(* IEC 61131-3 sources: plc-st-coding-agent/progress/evidence/f14_v14_remaining_20261113/jobs/custom_minimax-m27, 185 files *)

(* ---- public-easy-01.candidate_01.st ---- *)
(* ENGINEERING_CONTRACT
 * ============================================================================
 * State Machine: Automated Filling Line Control (6 states, sequential)
 * ============================================================================
 * | State      | Outputs Activated           | Retention    | Reset/Exit           |
 * |------------|-----------------------------|--------------|----------------------|
 * | IDLE       | none                        | -            | bottleSensor → CLEANING (PUB001) |
 * | CLEANING   | Pump_Motor:=TRUE            | hold until reset | cleaningConfirmButton → FILLING (PUB003) |
 * | FILLING    | Filling_Valve:=TRUE         | hold until reset | fillingConfirmButton → CAPPING (PUB003) |
 * | CAPPING    | Capping_Machine:=TRUE       | hold until reset | cappingConfirmButton → PACKING (PUB003) |
 * | PACKING    | Packing_Machine:=TRUE       | hold until reset | packingConfirmButton → COMPLETED (PUB005) |
 * | COMPLETED  | Completion_Light:=TRUE      | hold until reset | finishedButton → IDLE (PUB007) |
 * ============================================================================
 * Priority/Interlocks:
 *   - Physical direction rule: N/A (no opposite movements in this process)
 *   - Same-scan priority: outputs computed combinatorially from state, no priority
 *   - Button edge detection: R_TRIG on each confirm input to avoid repeat triggers
 *   - First scan behavior: outputs default to FALSE until first state transition
 *   - Boundary conditions: IDLE=0, COMPLETED=5 enum bounds, array indexing valid
 *   - Simultaneous buttons: not applicable (sequential process, one button per state)
 * ============================================================================
 * CONTRACT_RULES [{"kind": "hold_until_reset", "output": "Completion_Light", "set_input": "packingConfirmButton", "reset_input": "finishedButton"}]
 * ============================================================================
 *)

FUNCTION_BLOCK FillLineControl
VAR_INPUT
    bottleSensor          : BOOL;
    cleaningConfirmButton : BOOL;
    fillingConfirmButton  : BOOL;
    cappingConfirmButton  : BOOL;
    packingConfirmButton  : BOOL;
    finishedButton        : BOOL;
END_VAR
VAR_OUTPUT
    Pump_Motor      : BOOL;
    Filling_Valve   : BOOL;
    Capping_Machine : BOOL;
    Packing_Machine : BOOL;
    Completion_Light: BOOL;
END_VAR
VAR
    State        : UINT := 0;
    trg_bottle   : R_TRIG;
    trg_cleaning : R_TRIG;
    trg_filling  : R_TRIG;
    trg_capping  : R_TRIG;
    trg_packing  : R_TRIG;
    trg_finished : R_TRIG;
END_VAR

(* Constants for state identification *)
VAR CONSTANT
    STATE_IDLE      : UINT := 0;
    STATE_CLEANING  : UINT := 1;
    STATE_FILLING   : UINT := 2;
    STATE_CAPPING   : UINT := 3;
    STATE_PACKING   : UINT := 4;
    STATE_COMPLETED : UINT := 5;
END_VAR

(* Scan edge detectors *)
trg_bottle(CLK := bottleSensor);
trg_cleaning(CLK := cleaningConfirmButton);
trg_filling(CLK := fillingConfirmButton);
trg_capping(CLK := cappingConfirmButton);
trg_packing(CLK := packingConfirmButton);
trg_finished(CLK := finishedButton);

(* State machine transitions *)
CASE State OF
    STATE_IDLE:
        IF trg_bottle.Q THEN
            State := STATE_CLEANING;
        END_IF;

    STATE_CLEANING:
        IF trg_cleaning.Q THEN
            State := STATE_FILLING;
        END_IF;

    STATE_FILLING:
        IF trg_filling.Q THEN
            State := STATE_CAPPING;
        END_IF;

    STATE_CAPPING:
        IF trg_capping.Q THEN
            State := STATE_PACKING;
        END_IF;

    STATE_PACKING:
        IF trg_packing.Q THEN
            State := STATE_COMPLETED;
        END_IF;

    STATE_COMPLETED:
        IF trg_finished.Q THEN
            State := STATE_IDLE;
        END_IF;

END_CASE;

(* Output generation based on current state *)
Pump_Motor      := (State = STATE_CLEANING);
Filling_Valve   := (State = STATE_FILLING);
Capping_Machine := (State = STATE_CAPPING);
Packing_Machine := (State = STATE_PACKING);
Completion_Light:= (State = STATE_COMPLETED);

END_FUNCTION_BLOCK

(* ---- public-easy-01.raw_candidate_01.st ---- *)
(* ENGINEERING_CONTRACT
 * ============================================================================
 * State Machine: Automated Filling Line Control (6 states, sequential)
 * ============================================================================
 * | State      | Outputs Activated           | Retention    | Reset/Exit           |
 * |------------|-----------------------------|--------------|----------------------|
 * | IDLE       | none                        | -            | bottleSensor → CLEANING (PUB001) |
 * | CLEANING   | Pump_Motor:=TRUE            | hold until reset | cleaningConfirmButton → FILLING (PUB003) |
 * | FILLING    | Filling_Valve:=TRUE         | hold until reset | fillingConfirmButton → CAPPING (PUB003) |
 * | CAPPING    | Capping_Machine:=TRUE       | hold until reset | cappingConfirmButton → PACKING (PUB003) |
 * | PACKING    | Packing_Machine:=TRUE       | hold until reset | packingConfirmButton → COMPLETED (PUB005) |
 * | COMPLETED  | Completion_Light:=TRUE      | hold until reset | finishedButton → IDLE (PUB007) |
 * ============================================================================
 * Priority/Interlocks:
 *   - Physical direction rule: N/A (no opposite movements in this process)
 *   - Same-scan priority: outputs computed combinatorially from state, no priority
 *   - Button edge detection: R_TRIG on each confirm input to avoid repeat triggers
 *   - First scan behavior: outputs default to FALSE until first state transition
 *   - Boundary conditions: IDLE=0, COMPLETED=5 enum bounds, array indexing valid
 *   - Simultaneous buttons: not applicable (sequential process, one button per state)
 * ============================================================================
 * CONTRACT_RULES [{"kind": "hold_until_reset", "output": "Completion_Light", "set_input": "packingConfirmButton", "reset_input": "finishedButton"}]
 * ============================================================================
 *)

FUNCTION_BLOCK FillLineControl
VAR_INPUT
    bottleSensor          : BOOL;
    cleaningConfirmButton : BOOL;
    fillingConfirmButton  : BOOL;
    cappingConfirmButton  : BOOL;
    packingConfirmButton  : BOOL;
    finishedButton        : BOOL;
END_VAR
VAR_OUTPUT
    Pump_Motor      : BOOL;
    Filling_Valve   : BOOL;
    Capping_Machine : BOOL;
    Packing_Machine : BOOL;
    Completion_Light: BOOL;
END_VAR
VAR
    State        : UINT := 0;
    trg_bottle   : R_TRIG;
    trg_cleaning : R_TRIG;
    trg_filling  : R_TRIG;
    trg_capping  : R_TRIG;
    trg_packing  : R_TRIG;
    trg_finished : R_TRIG;
END_VAR

(* Constants for state identification *)
VAR CONSTANT
    STATE_IDLE      : UINT := 0;
    STATE_CLEANING  : UINT := 1;
    STATE_FILLING   : UINT := 2;
    STATE_CAPPING   : UINT := 3;
    STATE_PACKING   : UINT := 4;
    STATE_COMPLETED : UINT := 5;
END_VAR

(* Scan edge detectors *)
trg_bottle(CLK := bottleSensor);
trg_cleaning(CLK := cleaningConfirmButton);
trg_filling(CLK := fillingConfirmButton);
trg_capping(CLK := cappingConfirmButton);
trg_packing(CLK := packingConfirmButton);
trg_finished(CLK := finishedButton);

(* State machine transitions *)
CASE State OF
    STATE_IDLE:
        IF trg_bottle.Q THEN
            State := STATE_CLEANING;
        END_IF

    STATE_CLEANING:
        IF trg_cleaning.Q THEN
            State := STATE_FILLING;
        END_IF

    STATE_FILLING:
        IF trg_filling.Q THEN
            State := STATE_CAPPING;
        END_IF

    STATE_CAPPING:
        IF trg_capping.Q THEN
            State := STATE_PACKING;
        END_IF

    STATE_PACKING:
        IF trg_packing.Q THEN
            State := STATE_COMPLETED;
        END_IF

    STATE_COMPLETED:
        IF trg_finished.Q THEN
            State := STATE_IDLE;
        END_IF

END_CASE

(* Output generation based on current state *)
Pump_Motor      := (State = STATE_CLEANING);
Filling_Valve   := (State = STATE_FILLING);
Capping_Machine := (State = STATE_CAPPING);
Packing_Machine := (State = STATE_PACKING);
Completion_Light:= (State = STATE_COMPLETED);

END_FUNCTION_BLOCK

(* ---- public-easy-02.candidate_01.st ---- *)
FUNCTION_BLOCK FB_DualWordEdgeDetection
VAR_INPUT
    value : DWORD;
END_VAR

VAR_OUTPUT
    hasChanged       : BOOL;
    hasRisingEdges   : BOOL;
    risingBits       : DWORD;
    noOfRisingBits   : USINT;
    hasFallingEdges  : BOOL;
    fallingBits      : DWORD;
    noOfFallingBits  : USINT;
END_VAR

VAR
    prevValue : DWORD;
END_VAR

// ENGINEERING_CONTRACT:
// Outputs: hasChanged, hasRisingEdges, hasFallingEdges, risingBits, fallingBits, noOfRisingBits, noOfFallingBits
// Retention: All outputs retain their computed values across scans until recomputed.
// Reset: No explicit reset input defined; prevValue initializes to zero on first scan.
// Edge Detection: risingBits = value & ~prevValue; fallingBits = ~value & prevValue
// Counting: Iterates all 32 bits of risingBits/fallingBits to compute USINT counts.
// hasChanged = (value <> prevValue); hasRisingEdges = (risingBits <> 0); hasFallingEdges = (fallingBits <> 0)
// PUB001: Input value is DWORD; outputs report per-scan edge events.
// CONTRACT_RULES [{"kind": "hold_until_reset", "output": "risingBits", "set_input": "value", "reset_input": null}, {"kind": "hold_until_reset", "output": "fallingBits", "set_input": "value", "reset_input": null}, {"kind": "hold_until_reset", "output": "noOfRisingBits", "set_input": "value", "reset_input": null}, {"kind": "hold_until_reset", "output": "noOfFallingBits", "set_input": "value", "reset_input": null}]

risingBits  := value AND (NOT prevValue);
fallingBits := (NOT value) AND prevValue;

hasChanged      := (value <> prevValue);
hasRisingEdges  := (risingBits <> 16#00000000);
hasFallingEdges := (fallingBits <> 16#00000000);

noOfRisingBits  := 0;
noOfFallingBits := 0;

FOR i := 0 TO 31 DO
    IF (risingBits AND SHL(16#00000001, i)) <> 16#00000000 THEN
        noOfRisingBits := noOfRisingBits + 1;
    END_IF;

    IF (fallingBits AND SHL(16#00000001, i)) <> 16#00000000 THEN
        noOfFallingBits := noOfFallingBits + 1;
    END_IF;
END_FOR;

prevValue := value;

END_FUNCTION_BLOCK

(* ---- public-easy-02.candidate_02.st ---- *)
FUNCTION_BLOCK FB_DualWordEdgeDetection
VAR_INPUT
    value : DWORD;
END_VAR

VAR_OUTPUT
    hasChanged       : BOOL;
    hasRisingEdges   : BOOL;
    risingBits       : DWORD;
    noOfRisingBits   : USINT;
    hasFallingEdges  : BOOL;
    fallingBits      : DWORD;
    noOfFallingBits  : USINT;
END_VAR

VAR
    prevValue : DWORD;
    i         : UINT;
END_VAR

// ENGINEERING_CONTRACT:
// Outputs: hasChanged, hasRisingEdges, hasFallingEdges, risingBits, fallingBits, noOfRisingBits, noOfFallingBits
// Retention: All outputs retain their computed values across scans until recomputed.
// Reset: No explicit reset input defined; prevValue initializes to zero on first scan.
// Edge Detection: risingBits = value & ~prevValue; fallingBits = ~value & prevValue
// Counting: Iterates all 32 bits of risingBits/fallingBits to compute USINT counts.
// hasChanged = (value <> prevValue); hasRisingEdges = (risingBits <> 0); hasFallingEdges = (fallingBits <> 0)
// PUB001: Input value is DWORD; outputs report per-scan edge events.
// CONTRACT_RULES [{"kind": "hold_until_reset", "output": "risingBits", "set_input": "value", "reset_input": null}, {"kind": "hold_until_reset", "output": "fallingBits", "set_input": "value", "reset_input": null}, {"kind": "hold_until_reset", "output": "noOfRisingBits", "set_input": "value", "reset_input": null}, {"kind": "hold_until_reset", "output": "noOfFallingBits", "set_input": "value", "reset_input": null}]

risingBits  := value AND (NOT prevValue);
fallingBits := (NOT value) AND prevValue;

hasChanged      := (value <> prevValue);
hasRisingEdges  := (risingBits <> 16#00000000);
hasFallingEdges := (fallingBits <> 16#00000000);

noOfRisingBits  := 0;
noOfFallingBits := 0;

FOR i := 0 TO 31 DO
    IF (risingBits AND SHL(16#00000001, i)) <> 16#00000000 THEN
        noOfRisingBits := noOfRisingBits + 1;
    END_IF;

    IF (fallingBits AND SHL(16#00000001, i)) <> 16#00000000 THEN
        noOfFallingBits := noOfFallingBits + 1;
    END_IF;
END_FOR;

prevValue := value;

END_FUNCTION_BLOCK

(* ---- public-easy-02.patch_base_02.st ---- *)
FUNCTION_BLOCK FB_DualWordEdgeDetection
VAR_INPUT
    value : DWORD;
END_VAR

VAR_OUTPUT
    hasChanged       : BOOL;
    hasRisingEdges   : BOOL;
    risingBits       : DWORD;
    noOfRisingBits   : USINT;
    hasFallingEdges  : BOOL;
    fallingBits      : DWORD;
    noOfFallingBits  : USINT;
END_VAR

VAR
    prevValue : DWORD;
END_VAR

// ENGINEERING_CONTRACT:
// Outputs: hasChanged, hasRisingEdges, hasFallingEdges, risingBits, fallingBits, noOfRisingBits, noOfFallingBits
// Retention: All outputs retain their computed values across scans until recomputed.
// Reset: No explicit reset input defined; prevValue initializes to zero on first scan.
// Edge Detection: risingBits = value & ~prevValue; fallingBits = ~value & prevValue
// Counting: Iterates all 32 bits of risingBits/fallingBits to compute USINT counts.
// hasChanged = (value <> prevValue); hasRisingEdges = (risingBits <> 0); hasFallingEdges = (fallingBits <> 0)
// PUB001: Input value is DWORD; outputs report per-scan edge events.
// CONTRACT_RULES [{"kind": "hold_until_reset", "output": "risingBits", "set_input": "value", "reset_input": null}, {"kind": "hold_until_reset", "output": "fallingBits", "set_input": "value", "reset_input": null}, {"kind": "hold_until_reset", "output": "noOfRisingBits", "set_input": "value", "reset_input": null}, {"kind": "hold_until_reset", "output": "noOfFallingBits", "set_input": "value", "reset_input": null}]

risingBits  := value AND (NOT prevValue);
fallingBits := (NOT value) AND prevValue;

hasChanged      := (value <> prevValue);
hasRisingEdges  := (risingBits <> 16#00000000);
hasFallingEdges := (fallingBits <> 16#00000000);

noOfRisingBits  := 0;
noOfFallingBits := 0;

FOR i := 0 TO 31 DO
    IF (risingBits AND SHL(16#00000001, i)) <> 16#00000000 THEN
        noOfRisingBits := noOfRisingBits + 1;
    END_IF;

    IF (fallingBits AND SHL(16#00000001, i)) <> 16#00000000 THEN
        noOfFallingBits := noOfFallingBits + 1;
    END_IF;
END_FOR;

prevValue := value;

END_FUNCTION_BLOCK

(* ---- public-easy-02.raw_candidate_01.st ---- *)
FUNCTION_BLOCK FB_DualWordEdgeDetection
VAR_INPUT
    value : DWORD;
END_VAR

VAR_OUTPUT
    hasChanged       : BOOL;
    hasRisingEdges   : BOOL;
    risingBits       : DWORD;
    noOfRisingBits   : USINT;
    hasFallingEdges  : BOOL;
    fallingBits      : DWORD;
    noOfFallingBits  : USINT;
END_VAR

VAR
    prevValue : DWORD;
END_VAR

// ENGINEERING_CONTRACT:
// Outputs: hasChanged, hasRisingEdges, hasFallingEdges, risingBits, fallingBits, noOfRisingBits, noOfFallingBits
// Retention: All outputs retain their computed values across scans until recomputed.
// Reset: No explicit reset input defined; prevValue initializes to zero on first scan.
// Edge Detection: risingBits = value & ~prevValue; fallingBits = ~value & prevValue
// Counting: Iterates all 32 bits of risingBits/fallingBits to compute USINT counts.
// hasChanged = (value <> prevValue); hasRisingEdges = (risingBits <> 0); hasFallingEdges = (fallingBits <> 0)
// PUB001: Input value is DWORD; outputs report per-scan edge events.
// CONTRACT_RULES [{"kind": "hold_until_reset", "output": "risingBits", "set_input": "value", "reset_input": null}, {"kind": "hold_until_reset", "output": "fallingBits", "set_input": "value", "reset_input": null}, {"kind": "hold_until_reset", "output": "noOfRisingBits", "set_input": "value", "reset_input": null}, {"kind": "hold_until_reset", "output": "noOfFallingBits", "set_input": "value", "reset_input": null}]

risingBits  := value AND (NOT prevValue);
fallingBits := (NOT value) AND prevValue;

hasChanged      := (value <> prevValue);
hasRisingEdges  := (risingBits <> 16#00000000);
hasFallingEdges := (fallingBits <> 16#00000000);

noOfRisingBits  := 0;
noOfFallingBits := 0;

FOR i := 0 TO 31 DO
    IF (risingBits AND SHL(16#00000001, i)) <> 16#00000000 THEN
        noOfRisingBits := noOfRisingBits + 1;
    END_IF;

    IF (fallingBits AND SHL(16#00000001, i)) <> 16#00000000 THEN
        noOfFallingBits := noOfFallingBits + 1;
    END_IF;
END_FOR;

prevValue := value;

END_FUNCTION_BLOCK

(* ---- public-easy-02.raw_candidate_02.st ---- *)
FUNCTION_BLOCK FB_DualWordEdgeDetection
VAR_INPUT
    value : DWORD;
END_VAR

VAR_OUTPUT
    hasChanged       : BOOL;
    hasRisingEdges   : BOOL;
    risingBits       : DWORD;
    noOfRisingBits   : USINT;
    hasFallingEdges  : BOOL;
    fallingBits      : DWORD;
    noOfFallingBits  : USINT;
END_VAR

VAR
    prevValue : DWORD;
    i         : UINT;
END_VAR

// ENGINEERING_CONTRACT:
// Outputs: hasChanged, hasRisingEdges, hasFallingEdges, risingBits, fallingBits, noOfRisingBits, noOfFallingBits
// Retention: All outputs retain their computed values across scans until recomputed.
// Reset: No explicit reset input defined; prevValue initializes to zero on first scan.
// Edge Detection: risingBits = value & ~prevValue; fallingBits = ~value & prevValue
// Counting: Iterates all 32 bits of risingBits/fallingBits to compute USINT counts.
// hasChanged = (value <> prevValue); hasRisingEdges = (risingBits <> 0); hasFallingEdges = (fallingBits <> 0)
// PUB001: Input value is DWORD; outputs report per-scan edge events.
// CONTRACT_RULES [{"kind": "hold_until_reset", "output": "risingBits", "set_input": "value", "reset_input": null}, {"kind": "hold_until_reset", "output": "fallingBits", "set_input": "value", "reset_input": null}, {"kind": "hold_until_reset", "output": "noOfRisingBits", "set_input": "value", "reset_input": null}, {"kind": "hold_until_reset", "output": "noOfFallingBits", "set_input": "value", "reset_input": null}]

risingBits  := value AND (NOT prevValue);
fallingBits := (NOT value) AND prevValue;

hasChanged      := (value <> prevValue);
hasRisingEdges  := (risingBits <> 16#00000000);
hasFallingEdges := (fallingBits <> 16#00000000);

noOfRisingBits  := 0;
noOfFallingBits := 0;

FOR i := 0 TO 31 DO
    IF (risingBits AND SHL(16#00000001, i)) <> 16#00000000 THEN
        noOfRisingBits := noOfRisingBits + 1;
    END_IF;

    IF (fallingBits AND SHL(16#00000001, i)) <> 16#00000000 THEN
        noOfFallingBits := noOfFallingBits + 1;
    END_IF;
END_FOR;

prevValue := value;

END_FUNCTION_BLOCK

(* ---- public-easy-03.candidate_01.st ---- *)
FUNCTION_BLOCK AlarmHysteresis
VAR_INPUT
    Value      : REAL;
    hiLevel    : REAL;
    loLevel    : REAL;
    hystWindow : REAL;
END_VAR
VAR_OUTPUT
    hiAlarm : BOOL;
    loAlarm : BOOL;
    error   : BOOL;
    status  : WORD;
END_VAR
VAR
    tmp_range : REAL;
END_VAR

(* ENGINEERING_CONTRACT
| Output   | Activation                          | Retention        | Reset/Deactivation                  | Same-scan | Units/Bounds           |
|----------|-------------------------------------|------------------|-------------------------------------|-----------|------------------------|
| hiAlarm  | Value > hiLevel                     | hold             | Value < hiLevel - hystWindow        | -         | PUB001, hysteresis     |
| loAlarm  | Value < loLevel                     | hold             | Value > loLevel + hystWindow        | -         | PUB001, hysteresis     |
| error    | loLevel >= hiLevel                  | hold_until_reset | -                                   | priority  | PUB002, 16#8001        |
| error    | hystWindow >= (hiLevel - loLevel)   | hold_until_reset | -                                   | priority  | PUB003, 16#8002        |
| status   | set on error                        | retain           | -                                   | -         | PUB002/PUB003, WORD    |

Priority: Error checks execute before alarm logic; on error, status is set and block exits early.
Retention: hiAlarm/loAlarm are latching (PUB001); error is latching until explicit reset (not specified).
Boundary: Strict > and < comparisons; hystWindow is REAL; range = hiLevel - loLevel.
*)

(* CONTRACT_RULES [] *)

tmp_range := hiLevel - loLevel;

error := FALSE;
status := 16#0000;

IF loLevel >= hiLevel THEN
    error := TRUE;
    status := 16#8001;
    RETURN;
END_IF;

IF hystWindow >= tmp_range THEN
    error := TRUE;
    status := 16#8002;
    RETURN;
END_IF;

IF Value > hiLevel THEN
    hiAlarm := TRUE;
ELSIF Value < (hiLevel - hystWindow) THEN
    hiAlarm := FALSE;
END_IF;

IF Value < loLevel THEN
    loAlarm := TRUE;
ELSIF Value > (loLevel + hystWindow) THEN
    loAlarm := FALSE;
END_IF;

END_FUNCTION_BLOCK

(* ---- public-easy-03.raw_candidate_01.st ---- *)
FUNCTION_BLOCK AlarmHysteresis
VAR_INPUT
    Value      : REAL;
    hiLevel    : REAL;
    loLevel    : REAL;
    hystWindow : REAL;
END_VAR
VAR_OUTPUT
    hiAlarm : BOOL;
    loAlarm : BOOL;
    error   : BOOL;
    status  : WORD;
END_VAR
VAR
    tmp_range : REAL;
END_VAR

(* ENGINEERING_CONTRACT
| Output   | Activation                          | Retention        | Reset/Deactivation                  | Same-scan | Units/Bounds           |
|----------|-------------------------------------|------------------|-------------------------------------|-----------|------------------------|
| hiAlarm  | Value > hiLevel                     | hold             | Value < hiLevel - hystWindow        | -         | PUB001, hysteresis     |
| loAlarm  | Value < loLevel                     | hold             | Value > loLevel + hystWindow        | -         | PUB001, hysteresis     |
| error    | loLevel >= hiLevel                  | hold_until_reset | -                                   | priority  | PUB002, 16#8001        |
| error    | hystWindow >= (hiLevel - loLevel)   | hold_until_reset | -                                   | priority  | PUB003, 16#8002        |
| status   | set on error                        | retain           | -                                   | -         | PUB002/PUB003, WORD    |

Priority: Error checks execute before alarm logic; on error, status is set and block exits early.
Retention: hiAlarm/loAlarm are latching (PUB001); error is latching until explicit reset (not specified).
Boundary: Strict > and < comparisons; hystWindow is REAL; range = hiLevel - loLevel.
*)

(* CONTRACT_RULES [] *)

tmp_range := hiLevel - loLevel;

error := FALSE;
status := 16#0000;

IF loLevel >= hiLevel THEN
    error := TRUE;
    status := 16#8001;
    RETURN;
END_IF

IF hystWindow >= tmp_range THEN
    error := TRUE;
    status := 16#8002;
    RETURN;
END_IF

IF Value > hiLevel THEN
    hiAlarm := TRUE;
ELSIF Value < (hiLevel - hystWindow) THEN
    hiAlarm := FALSE;
END_IF

IF Value < loLevel THEN
    loAlarm := TRUE;
ELSIF Value > (loLevel + hystWindow) THEN
    loAlarm := FALSE;
END_IF

END_FUNCTION_BLOCK

(* ---- public-easy-04.candidate_01.st ---- *)
(* ENGINEERING_CONTRACT:
1. VFD_RUN: Activation=debounced_viscosity AND PASTE_E_STOP_NC; Retention=held continuously while both inputs valid; Reset=immediate on E_STOP_NC=FALSE or viscosity invalid; Same-scan priority=evaluate after debounce state is finalized.
2. Viscosity debounce (TON): Activation=starts when VISCOSITY_OK=TRUE; Condition=VISCOSITY_OK must remain TRUE for DebounceTime; Reset=immediately when VISCOSITY_OK=FALSE or E_STOP_NC=FALSE (clears incomplete timing).
3. PUMP_RUNTIME_ACC: Activation=accumulates CycleTime each scan when VFD_RUN=TRUE; Retention=preserved when VFD_RUN=FALSE; Reset=none except power-up to 0 LTIME; Units=LTIME nanoseconds.
4. PUMP_MAINT_DUE: Activation=acc >= 500 hours (1,800,000,000 ms as LTIME); Retention=latched TRUE until power cycle; Reset=power cycle only; No effect on VFD_RUN or safety permissive.
5. Power-up: VFD_RUN=FALSE, PUMP_RUNTIME_ACC=0 LTIME, PUMP_MAINT_DUE=FALSE.
*)

(* CONTRACT_RULES: [{"kind": "hold_until_reset", "output": "PUMP_MAINT_DUE", "set_input": null, "reset_input": null}] *)

FUNCTION_BLOCK JamPumpControl
VAR_OUTPUT
    VFD_RUN            : BOOL  := FALSE;
    PUMP_MAINT_DUE     : BOOL  := FALSE;
    PUMP_RUNTIME_ACC   : LTIME := LTIME#0s;
END_VAR
VAR_INPUT
    VISCOSITY_OK       : BOOL;
    PASTE_E_STOP_NC    : BOOL;
    DebounceTime       : TIME;
    CycleTime          : TIME;
END_VAR
VAR
    tmp_debounce_ok    : BOOL := FALSE;
    debounce_timer     : TON;
END_VAR

    // Clear debounce timer immediately when emergency stop is released
    IF NOT PASTE_E_STOP_NC THEN
        debounce_timer(IN := FALSE, PT := DebounceTime);
        tmp_debounce_ok := FALSE;
    ELSE
        // Invalidate debounce immediately when viscosity signal drops
        IF NOT VISCOSITY_OK THEN
            debounce_timer(IN := FALSE, PT := DebounceTime);
            tmp_debounce_ok := FALSE;
        ELSE
            // Start or continue debounce timing while viscosity is valid
            debounce_timer(IN := TRUE, PT := DebounceTime);
            tmp_debounce_ok := debounce_timer.Q;
        END_IF;
    END_IF;

    // Set maintenance flag when runtime reaches 500 hours (latching)
    IF PUMP_RUNTIME_ACC >= LTIME#500h THEN
        PUMP_MAINT_DUE := TRUE;
    END_IF;

    // VFD run command: requires valid debounced viscosity AND no emergency stop
    VFD_RUN := tmp_debounce_ok AND PASTE_E_STOP_NC;

    // Accumulate runtime only while pump is running
    IF VFD_RUN THEN
        PUMP_RUNTIME_ACC := PUMP_RUNTIME_ACC + TO_LTIME(CycleTime);
    END_IF;

END_FUNCTION_BLOCK

(* ---- public-easy-04.patch_base_02.st ---- *)
(* ENGINEERING_CONTRACT:
1. VFD_RUN: Activation=debounced_viscosity AND PASTE_E_STOP_NC; Retention=held continuously while both inputs valid; Reset=immediate on E_STOP_NC=FALSE or viscosity invalid; Same-scan priority=evaluate after debounce state is finalized.
2. Viscosity debounce (TON): Activation=starts when VISCOSITY_OK=TRUE; Condition=VISCOSITY_OK must remain TRUE for DebounceTime; Reset=immediately when VISCOSITY_OK=FALSE or E_STOP_NC=FALSE (clears incomplete timing).
3. PUMP_RUNTIME_ACC: Activation=accumulates CycleTime each scan when VFD_RUN=TRUE; Retention=preserved when VFD_RUN=FALSE; Reset=none except power-up to 0 LTIME; Units=LTIME nanoseconds.
4. PUMP_MAINT_DUE: Activation=acc >= 500 hours (1,800,000,000 ms as LTIME); Retention=latched TRUE until power cycle; Reset=power cycle only; No effect on VFD_RUN or safety permissive.
5. Power-up: VFD_RUN=FALSE, PUMP_RUNTIME_ACC=0 LTIME, PUMP_MAINT_DUE=FALSE.
*)

(* CONTRACT_RULES: [{"kind": "hold_until_reset", "output": "PUMP_MAINT_DUE", "set_input": null, "reset_input": null}] *)

FUNCTION_BLOCK JamPumpControl
VAR_OUTPUT
    VFD_RUN            : BOOL  := FALSE;
    PUMP_MAINT_DUE     : BOOL  := FALSE;
    PUMP_RUNTIME_ACC   : LTIME := LTIME#0s;
END_VAR
VAR_INPUT
    VISCOSITY_OK       : BOOL;
    PASTE_E_STOP_NC    : BOOL;
    DebounceTime       : TIME;
    CycleTime          : TIME;
END_VAR
VAR
    tmp_debounce_ok    : BOOL := FALSE;
    debounce_timer     : TON;
END_VAR

    // Clear debounce timer immediately when emergency stop is released
    IF NOT PASTE_E_STOP_NC THEN
        debounce_timer(IN := FALSE, PT := DebounceTime);
        tmp_debounce_ok := FALSE;
    ELSE
        // Invalidate debounce immediately when viscosity signal drops
        IF NOT VISCOSITY_OK THEN
            debounce_timer(IN := FALSE, PT := DebounceTime);
            tmp_debounce_ok := FALSE;
        ELSE
            // Start or continue debounce timing while viscosity is valid
            debounce_timer(IN := TRUE, PT := DebounceTime);
            tmp_debounce_ok := debounce_timer.Q;
        END_IF;
    END_IF;

    // Set maintenance flag when runtime reaches 500 hours (latching)
    IF PUMP_RUNTIME_ACC >= LTIME#500h THEN
        PUMP_MAINT_DUE := TRUE;
    END_IF;

    // VFD run command: requires valid debounced viscosity AND no emergency stop
    VFD_RUN := tmp_debounce_ok AND PASTE_E_STOP_NC;

    // Accumulate runtime only while pump is running
    IF VFD_RUN THEN
        PUMP_RUNTIME_ACC := PUMP_RUNTIME_ACC + TO_LTIME(CycleTime);
    END_IF;

END_FUNCTION_BLOCK

(* ---- public-easy-04.patch_base_03.st ---- *)
(* ENGINEERING_CONTRACT:
1. VFD_RUN: Activation=debounced_viscosity AND PASTE_E_STOP_NC; Retention=held continuously while both inputs valid; Reset=immediate on E_STOP_NC=FALSE or viscosity invalid; Same-scan priority=evaluate after debounce state is finalized.
2. Viscosity debounce (TON): Activation=starts when VISCOSITY_OK=TRUE; Condition=VISCOSITY_OK must remain TRUE for DebounceTime; Reset=immediately when VISCOSITY_OK=FALSE or E_STOP_NC=FALSE (clears incomplete timing).
3. PUMP_RUNTIME_ACC: Activation=accumulates CycleTime each scan when VFD_RUN=TRUE; Retention=preserved when VFD_RUN=FALSE; Reset=none except power-up to 0 LTIME; Units=LTIME nanoseconds.
4. PUMP_MAINT_DUE: Activation=acc >= 500 hours (1,800,000,000 ms as LTIME); Retention=latched TRUE until power cycle; Reset=power cycle only; No effect on VFD_RUN or safety permissive.
5. Power-up: VFD_RUN=FALSE, PUMP_RUNTIME_ACC=0 LTIME, PUMP_MAINT_DUE=FALSE.
*)

(* CONTRACT_RULES: [{"kind": "hold_until_reset", "output": "PUMP_MAINT_DUE", "set_input": null, "reset_input": null}] *)

FUNCTION_BLOCK JamPumpControl
VAR_OUTPUT
    VFD_RUN            : BOOL  := FALSE;
    PUMP_MAINT_DUE     : BOOL  := FALSE;
    PUMP_RUNTIME_ACC   : LTIME := LTIME#0s;
END_VAR
VAR_INPUT
    VISCOSITY_OK       : BOOL;
    PASTE_E_STOP_NC    : BOOL;
    DebounceTime       : TIME;
    CycleTime          : TIME;
END_VAR
VAR
    tmp_debounce_ok    : BOOL := FALSE;
    debounce_timer     : TON;
END_VAR

    // Clear debounce timer immediately when emergency stop is released
    IF NOT PASTE_E_STOP_NC THEN
        debounce_timer(IN := FALSE, PT := DebounceTime);
        tmp_debounce_ok := FALSE;
    ELSE
        // Invalidate debounce immediately when viscosity signal drops
        IF NOT VISCOSITY_OK THEN
            debounce_timer(IN := FALSE, PT := DebounceTime);
            tmp_debounce_ok := FALSE;
        ELSE
            // Start or continue debounce timing while viscosity is valid
            debounce_timer(IN := TRUE, PT := DebounceTime);
            tmp_debounce_ok := debounce_timer.Q;
        END_IF;
    END_IF;

    // Set maintenance flag when runtime reaches 500 hours (latching)
    IF PUMP_RUNTIME_ACC >= LTIME#500h THEN
        PUMP_MAINT_DUE := TRUE;
    END_IF;

    // VFD run command: requires valid debounced viscosity AND no emergency stop
    VFD_RUN := tmp_debounce_ok AND PASTE_E_STOP_NC;

    // Accumulate runtime only while pump is running
    IF VFD_RUN THEN
        PUMP_RUNTIME_ACC := PUMP_RUNTIME_ACC + TO_LTIME(CycleTime);
    END_IF;

END_FUNCTION_BLOCK

(* ---- public-easy-04.raw_candidate_01.st ---- *)
(* ENGINEERING_CONTRACT:
1. VFD_RUN: Activation=debounced_viscosity AND PASTE_E_STOP_NC; Retention=held continuously while both inputs valid; Reset=immediate on E_STOP_NC=FALSE or viscosity invalid; Same-scan priority=evaluate after debounce state is finalized.
2. Viscosity debounce (TON): Activation=starts when VISCOSITY_OK=TRUE; Condition=VISCOSITY_OK must remain TRUE for DebounceTime; Reset=immediately when VISCOSITY_OK=FALSE or E_STOP_NC=FALSE (clears incomplete timing).
3. PUMP_RUNTIME_ACC: Activation=accumulates CycleTime each scan when VFD_RUN=TRUE; Retention=preserved when VFD_RUN=FALSE; Reset=none except power-up to 0 LTIME; Units=LTIME nanoseconds.
4. PUMP_MAINT_DUE: Activation=acc >= 500 hours (1,800,000,000 ms as LTIME); Retention=latched TRUE until power cycle; Reset=power cycle only; No effect on VFD_RUN or safety permissive.
5. Power-up: VFD_RUN=FALSE, PUMP_RUNTIME_ACC=0 LTIME, PUMP_MAINT_DUE=FALSE.
*)

(* CONTRACT_RULES: [{"kind": "hold_until_reset", "output": "PUMP_MAINT_DUE", "set_input": null, "reset_input": null}] *)

FUNCTION_BLOCK JamPumpControl
VAR_OUTPUT
    VFD_RUN            : BOOL  := FALSE;
    PUMP_MAINT_DUE     : BOOL  := FALSE;
    PUMP_RUNTIME_ACC   : LTIME := LTIME#0s;
END_VAR
VAR_INPUT
    VISCOSITY_OK       : BOOL;
    PASTE_E_STOP_NC    : BOOL;
    DebounceTime       : TIME;
    CycleTime          : TIME;
END_VAR
VAR
    tmp_debounce_ok    : BOOL := FALSE;
    debounce_timer     : TON;
END_VAR

    // Clear debounce timer immediately when emergency stop is released
    IF NOT PASTE_E_STOP_NC THEN
        debounce_timer(IN := FALSE, PT := DebounceTime);
        tmp_debounce_ok := FALSE;
    ELSE
        // Invalidate debounce immediately when viscosity signal drops
        IF NOT VISCOSITY_OK THEN
            debounce_timer(IN := FALSE, PT := DebounceTime);
            tmp_debounce_ok := FALSE;
        ELSE
            // Start or continue debounce timing while viscosity is valid
            debounce_timer(IN := TRUE, PT := DebounceTime);
            tmp_debounce_ok := debounce_timer.Q;
        END_IF;
    END_IF;

    // Set maintenance flag when runtime reaches 500 hours (latching)
    IF PUMP_RUNTIME_ACC >= LTIME#500h THEN
        PUMP_MAINT_DUE := TRUE;
    END_IF;

    // VFD run command: requires valid debounced viscosity AND no emergency stop
    VFD_RUN := tmp_debounce_ok AND PASTE_E_STOP_NC;

    // Accumulate runtime only while pump is running
    IF VFD_RUN THEN
        PUMP_RUNTIME_ACC := PUMP_RUNTIME_ACC + TO_LTIME(CycleTime);
    END_IF;

END_FUNCTION_BLOCK

(* ---- public-easy-05.candidate_01.st ---- *)
FUNCTION_BLOCK WeldGapAlarm
(* ENGINEERING_CONTRACT
   =================================================================
   States & Retention (outputs per PUB001-PUB006):
   -----------------------------------------------------------------
   State: POWER_UP_INHIBIT (5s after power-up, no E-stop)
   - Weld_Soft_Start_Active := TRUE (activation: power-up entry)
   - Operator_Alert := FALSE (held, no alarm during inhibit)
   - Gap debounce does NOT accumulate (timer gated OFF)
   - Retention: held until 5s elapsed OR E-stop asserted
   -----------------------------------------------------------------
   State: NORMAL_MONITORING (after 5s inhibit, no E-stop)
   - Weld_Soft_Start_Active := FALSE (deactivated, no reset input)
   - Operator_Alert := TRUE only when DebounceTimer.Q = TRUE
     (activation: Gap_Exceeded TRUE for DebounceTime; retention:
      held until Gap_Exceeded FALSE OR E-stop asserted)
   - DebounceTimer enabled when Gap_Exceeded = TRUE; cleared when
     Gap_Exceeded = FALSE; no same-scan priority issue (TON called
     once with final enable state)
   - Reset: E-stop immediate reset, then return to POWER_UP_INHIBIT
   -----------------------------------------------------------------
   E-STOP PRIORITY (Weld_E_Stop_NC = FALSE):
   - Operator_Alert immediately FALSE (explicit reset per PUB004)
   - Incomplete debounce timing cleared (TON.ET reset via re-call
     with IN=FALSE when E-stop detected)
   - Weld_Soft_Start_Active := FALSE (inhibition cancelled)
   - Same-scan: evaluated before state logic; no race condition
   -----------------------------------------------------------------
   Units/Boundaries:
   - Power-up inhibit: 5s (T#5s), LTIME resolution
   - DebounceTime: caller-supplied TIME, must be positive (PUB003)
   - TON.Q activates at ET >= PT; ET saturates at PT
   - Direction conflicts: not applicable (no axis outputs)
   =================================================================
*)
VAR
    // Power-up initialization timer: 5-second inhibit period
    PowerUpTimer: TON;
    // Gap signal debounce timer during normal monitoring
    DebounceTimer: TON;
END_VAR

// E-STOP PRIORITY: Immediate deactivation per PUB004
// Evaluated first to ensure same-scan priority over state transitions
IF NOT Weld_E_Stop_NC THEN
    // Operator_Alert immediately FALSE
    Operator_Alert := FALSE;
    // Clear any incomplete debounce timing (re-call with IN=FALSE clears ET)
    DebounceTimer(IN := FALSE, PT := DebounceTime);
    // Cancel power-up inhibition (soft start no longer valid)
    Weld_Soft_Start_Active := FALSE;
    // Restart power-up timer on next rising edge of E-stop release
    PowerUpTimer(IN := FALSE, PT := T#5s);
ELSE
    // E-stop inactive (Weld_E_Stop_NC = TRUE): normal/state logic

    // Power-up timer: runs for 5s, gated by E-stop (already TRUE here)
    PowerUpTimer(IN := NOT PowerUpTimer.Q, PT := T#5s);

    // Determine current operating phase
    IF NOT PowerUpTimer.Q THEN
        // POWER_UP_INHIBIT state: 5-second initialization period
        // PUB001: Operator_Alert = FALSE during inhibit
        Operator_Alert := FALSE;
        // PUB002: Weld_Soft_Start_Active = TRUE during inhibit
        Weld_Soft_Start_Active := TRUE;
        // PUB003: Gap debounce time does NOT accumulate during inhibit
        // Timer not called, so no timing accumulation
    ELSE
        // NORMAL_MONITORING state: after 5-second inhibit completes
        // PUB002: Weld_Soft_Start_Active = FALSE after inhibit
        Weld_Soft_Start_Active := FALSE;

        // Debounce logic: accumulate time only when Gap_Exceeded = TRUE
        // When Gap_Exceeded = FALSE, timer resets (IN=FALSE clears ET)
        DebounceTimer(
            IN := Gap_Exceeded,
            PT := DebounceTime
        );

        // Operator_Alert activated after debounce completes (PUB003)
        // Retention: remains TRUE until Gap_Exceeded FALSE OR E-stop
        Operator_Alert := DebounceTimer.Q;
    END_IF;
END_IF;
END_FUNCTION_BLOCK

(* ---- public-easy-05.candidate_02.st ---- *)
FUNCTION_BLOCK WeldGapAlarm
(* ENGINEERING_CONTRACT
   =================================================================
   States & Retention (outputs per PUB001-PUB006):
   -----------------------------------------------------------------
   State: POWER_UP_INHIBIT (5s after power-up, no E-stop)
   - Weld_Soft_Start_Active := TRUE (activation: power-up entry)
   - Operator_Alert := FALSE (held, no alarm during inhibit)
   - Gap debounce does NOT accumulate (timer gated OFF)
   - Retention: held until 5s elapsed OR E-stop asserted
   -----------------------------------------------------------------
   State: NORMAL_MONITORING (after 5s inhibit, no E-stop)
   - Weld_Soft_Start_Active := FALSE (deactivated, no reset input)
   - Operator_Alert := TRUE only when DebounceTimer.Q = TRUE
     (activation: Gap_Exceeded TRUE for DebounceTime; retention:
      held until Gap_Exceeded FALSE OR E-stop asserted)
   - DebounceTimer enabled when Gap_Exceeded = TRUE; cleared when
     Gap_Exceeded = FALSE; no same-scan priority issue (TON called
     once with final enable state)
   - Reset: E-stop immediate reset, then return to POWER_UP_INHIBIT
   -----------------------------------------------------------------
   E-STOP PRIORITY (Weld_E_Stop_NC = FALSE):
   - Operator_Alert immediately FALSE (explicit reset per PUB004)
   - Incomplete debounce timing cleared (TON.ET reset via re-call
     with IN=FALSE when E-stop detected)
   - Weld_Soft_Start_Active := FALSE (inhibition cancelled)
   - Same-scan: evaluated before state logic; no race condition
   -----------------------------------------------------------------
   Units/Boundaries:
   - Power-up inhibit: 5s (T#5s), LTIME resolution
   - DebounceTime: caller-supplied TIME, must be positive (PUB003)
   - TON.Q activates at ET >= PT; ET saturates at PT
   - Direction conflicts: not applicable (no axis outputs)
   =================================================================
*)
VAR_INPUT
    Gap_Exceeded: BOOL;
    Weld_E_Stop_NC: BOOL;
    DebounceTime: TIME;
END_VAR

VAR_OUTPUT
    Operator_Alert: BOOL;
    Weld_Soft_Start_Active: BOOL;
END_VAR

VAR
    // Power-up initialization timer: 5-second inhibit period
    PowerUpTimer: TON;
    // Gap signal debounce timer during normal monitoring
    DebounceTimer: TON;
END_VAR

// E-STOP PRIORITY: Immediate deactivation per PUB004
// Evaluated first to ensure same-scan priority over state transitions
IF NOT Weld_E_Stop_NC THEN
    // Operator_Alert immediately FALSE
    Operator_Alert := FALSE;
    // Clear any incomplete debounce timing (re-call with IN=FALSE clears ET)
    DebounceTimer(IN := FALSE, PT := DebounceTime);
    // Cancel power-up inhibition (soft start no longer valid)
    Weld_Soft_Start_Active := FALSE;
    // Restart power-up timer on next rising edge of E-stop release
    PowerUpTimer(IN := FALSE, PT := T#5s);
ELSE
    // E-stop inactive (Weld_E_Stop_NC = TRUE): normal/state logic

    // Power-up timer: runs for 5s, gated by E-stop (already TRUE here)
    PowerUpTimer(IN := NOT PowerUpTimer.Q, PT := T#5s);

    // Determine current operating phase
    IF NOT PowerUpTimer.Q THEN
        // POWER_UP_INHIBIT state: 5-second initialization period
        // PUB001: Operator_Alert = FALSE during inhibit
        Operator_Alert := FALSE;
        // PUB002: Weld_Soft_Start_Active = TRUE during inhibit
        Weld_Soft_Start_Active := TRUE;
        // PUB003: Gap debounce time does NOT accumulate during inhibit
        // Timer not called, so no timing accumulation
    ELSE
        // NORMAL_MONITORING state: after 5-second inhibit completes
        // PUB002: Weld_Soft_Start_Active = FALSE after inhibit
        Weld_Soft_Start_Active := FALSE;

        // Debounce logic: accumulate time only when Gap_Exceeded = TRUE
        // When Gap_Exceeded = FALSE, timer resets (IN=FALSE clears ET)
        DebounceTimer(
            IN := Gap_Exceeded,
            PT := DebounceTime
        );

        // Operator_Alert activated after debounce completes (PUB003)
        // Retention: remains TRUE until Gap_Exceeded FALSE OR E-stop
        Operator_Alert := DebounceTimer.Q;
    END_IF;
END_IF;
END_FUNCTION_BLOCK

(* ---- public-easy-05.patch_base_02.st ---- *)
FUNCTION_BLOCK WeldGapAlarm
(* ENGINEERING_CONTRACT
   =================================================================
   States & Retention (outputs per PUB001-PUB006):
   -----------------------------------------------------------------
   State: POWER_UP_INHIBIT (5s after power-up, no E-stop)
   - Weld_Soft_Start_Active := TRUE (activation: power-up entry)
   - Operator_Alert := FALSE (held, no alarm during inhibit)
   - Gap debounce does NOT accumulate (timer gated OFF)
   - Retention: held until 5s elapsed OR E-stop asserted
   -----------------------------------------------------------------
   State: NORMAL_MONITORING (after 5s inhibit, no E-stop)
   - Weld_Soft_Start_Active := FALSE (deactivated, no reset input)
   - Operator_Alert := TRUE only when DebounceTimer.Q = TRUE
     (activation: Gap_Exceeded TRUE for DebounceTime; retention:
      held until Gap_Exceeded FALSE OR E-stop asserted)
   - DebounceTimer enabled when Gap_Exceeded = TRUE; cleared when
     Gap_Exceeded = FALSE; no same-scan priority issue (TON called
     once with final enable state)
   - Reset: E-stop immediate reset, then return to POWER_UP_INHIBIT
   -----------------------------------------------------------------
   E-STOP PRIORITY (Weld_E_Stop_NC = FALSE):
   - Operator_Alert immediately FALSE (explicit reset per PUB004)
   - Incomplete debounce timing cleared (TON.ET reset via re-call
     with IN=FALSE when E-stop detected)
   - Weld_Soft_Start_Active := FALSE (inhibition cancelled)
   - Same-scan: evaluated before state logic; no race condition
   -----------------------------------------------------------------
   Units/Boundaries:
   - Power-up inhibit: 5s (T#5s), LTIME resolution
   - DebounceTime: caller-supplied TIME, must be positive (PUB003)
   - TON.Q activates at ET >= PT; ET saturates at PT
   - Direction conflicts: not applicable (no axis outputs)
   =================================================================
*)
VAR
    // Power-up initialization timer: 5-second inhibit period
    PowerUpTimer: TON;
    // Gap signal debounce timer during normal monitoring
    DebounceTimer: TON;
END_VAR

// E-STOP PRIORITY: Immediate deactivation per PUB004
// Evaluated first to ensure same-scan priority over state transitions
IF NOT Weld_E_Stop_NC THEN
    // Operator_Alert immediately FALSE
    Operator_Alert := FALSE;
    // Clear any incomplete debounce timing (re-call with IN=FALSE clears ET)
    DebounceTimer(IN := FALSE, PT := DebounceTime);
    // Cancel power-up inhibition (soft start no longer valid)
    Weld_Soft_Start_Active := FALSE;
    // Restart power-up timer on next rising edge of E-stop release
    PowerUpTimer(IN := FALSE, PT := T#5s);
ELSE
    // E-stop inactive (Weld_E_Stop_NC = TRUE): normal/state logic

    // Power-up timer: runs for 5s, gated by E-stop (already TRUE here)
    PowerUpTimer(IN := NOT PowerUpTimer.Q, PT := T#5s);

    // Determine current operating phase
    IF NOT PowerUpTimer.Q THEN
        // POWER_UP_INHIBIT state: 5-second initialization period
        // PUB001: Operator_Alert = FALSE during inhibit
        Operator_Alert := FALSE;
        // PUB002: Weld_Soft_Start_Active = TRUE during inhibit
        Weld_Soft_Start_Active := TRUE;
        // PUB003: Gap debounce time does NOT accumulate during inhibit
        // Timer not called, so no timing accumulation
    ELSE
        // NORMAL_MONITORING state: after 5-second inhibit completes
        // PUB002: Weld_Soft_Start_Active = FALSE after inhibit
        Weld_Soft_Start_Active := FALSE;

        // Debounce logic: accumulate time only when Gap_Exceeded = TRUE
        // When Gap_Exceeded = FALSE, timer resets (IN=FALSE clears ET)
        DebounceTimer(
            IN := Gap_Exceeded,
            PT := DebounceTime
        );

        // Operator_Alert activated after debounce completes (PUB003)
        // Retention: remains TRUE until Gap_Exceeded FALSE OR E-stop
        Operator_Alert := DebounceTimer.Q;
    END_IF;
END_IF;
END_FUNCTION_BLOCK

(* ---- public-easy-05.patch_base_03.st ---- *)
FUNCTION_BLOCK WeldGapAlarm
(* ENGINEERING_CONTRACT
   =================================================================
   States & Retention (outputs per PUB001-PUB006):
   -----------------------------------------------------------------
   State: POWER_UP_INHIBIT (5s after power-up, no E-stop)
   - Weld_Soft_Start_Active := TRUE (activation: power-up entry)
   - Operator_Alert := FALSE (held, no alarm during inhibit)
   - Gap debounce does NOT accumulate (timer gated OFF)
   - Retention: held until 5s elapsed OR E-stop asserted
   -----------------------------------------------------------------
   State: NORMAL_MONITORING (after 5s inhibit, no E-stop)
   - Weld_Soft_Start_Active := FALSE (deactivated, no reset input)
   - Operator_Alert := TRUE only when DebounceTimer.Q = TRUE
     (activation: Gap_Exceeded TRUE for DebounceTime; retention:
      held until Gap_Exceeded FALSE OR E-stop asserted)
   - DebounceTimer enabled when Gap_Exceeded = TRUE; cleared when
     Gap_Exceeded = FALSE; no same-scan priority issue (TON called
     once with final enable state)
   - Reset: E-stop immediate reset, then return to POWER_UP_INHIBIT
   -----------------------------------------------------------------
   E-STOP PRIORITY (Weld_E_Stop_NC = FALSE):
   - Operator_Alert immediately FALSE (explicit reset per PUB004)
   - Incomplete debounce timing cleared (TON.ET reset via re-call
     with IN=FALSE when E-stop detected)
   - Weld_Soft_Start_Active := FALSE (inhibition cancelled)
   - Same-scan: evaluated before state logic; no race condition
   -----------------------------------------------------------------
   Units/Boundaries:
   - Power-up inhibit: 5s (T#5s), LTIME resolution
   - DebounceTime: caller-supplied TIME, must be positive (PUB003)
   - TON.Q activates at ET >= PT; ET saturates at PT
   - Direction conflicts: not applicable (no axis outputs)
   =================================================================
*)
VAR_INPUT
    Gap_Exceeded: BOOL;
    Weld_E_Stop_NC: BOOL;
    DebounceTime: TIME;
END_VAR

VAR_OUTPUT
    Operator_Alert: BOOL;
    Weld_Soft_Start_Active: BOOL;
END_VAR

VAR
    // Power-up initialization timer: 5-second inhibit period
    PowerUpTimer: TON;
    // Gap signal debounce timer during normal monitoring
    DebounceTimer: TON;
END_VAR

// E-STOP PRIORITY: Immediate deactivation per PUB004
// Evaluated first to ensure same-scan priority over state transitions
IF NOT Weld_E_Stop_NC THEN
    // Operator_Alert immediately FALSE
    Operator_Alert := FALSE;
    // Clear any incomplete debounce timing (re-call with IN=FALSE clears ET)
    DebounceTimer(IN := FALSE, PT := DebounceTime);
    // Cancel power-up inhibition (soft start no longer valid)
    Weld_Soft_Start_Active := FALSE;
    // Restart power-up timer on next rising edge of E-stop release
    PowerUpTimer(IN := FALSE, PT := T#5s);
ELSE
    // E-stop inactive (Weld_E_Stop_NC = TRUE): normal/state logic

    // Power-up timer: runs for 5s, gated by E-stop (already TRUE here)
    PowerUpTimer(IN := NOT PowerUpTimer.Q, PT := T#5s);

    // Determine current operating phase
    IF NOT PowerUpTimer.Q THEN
        // POWER_UP_INHIBIT state: 5-second initialization period
        // PUB001: Operator_Alert = FALSE during inhibit
        Operator_Alert := FALSE;
        // PUB002: Weld_Soft_Start_Active = TRUE during inhibit
        Weld_Soft_Start_Active := TRUE;
        // PUB003: Gap debounce time does NOT accumulate during inhibit
        // Timer not called, so no timing accumulation
    ELSE
        // NORMAL_MONITORING state: after 5-second inhibit completes
        // PUB002: Weld_Soft_Start_Active = FALSE after inhibit
        Weld_Soft_Start_Active := FALSE;

        // Debounce logic: accumulate time only when Gap_Exceeded = TRUE
        // When Gap_Exceeded = FALSE, timer resets (IN=FALSE clears ET)
        DebounceTimer(
            IN := Gap_Exceeded,
            PT := DebounceTime
        );

        // Operator_Alert activated after debounce completes (PUB003)
        // Retention: remains TRUE until Gap_Exceeded FALSE OR E-stop
        Operator_Alert := DebounceTimer.Q;
    END_IF;
END_IF;
END_FUNCTION_BLOCK

(* ---- public-easy-05.patch_base_04.st ---- *)
FUNCTION_BLOCK WeldGapAlarm
(* ENGINEERING_CONTRACT
   =================================================================
   States & Retention (outputs per PUB001-PUB006):
   -----------------------------------------------------------------
   State: POWER_UP_INHIBIT (5s after power-up, no E-stop)
   - Weld_Soft_Start_Active := TRUE (activation: power-up entry)
   - Operator_Alert := FALSE (held, no alarm during inhibit)
   - Gap debounce does NOT accumulate (timer gated OFF)
   - Retention: held until 5s elapsed OR E-stop asserted
   -----------------------------------------------------------------
   State: NORMAL_MONITORING (after 5s inhibit, no E-stop)
   - Weld_Soft_Start_Active := FALSE (deactivated, no reset input)
   - Operator_Alert := TRUE only when DebounceTimer.Q = TRUE
     (activation: Gap_Exceeded TRUE for DebounceTime; retention:
      held until Gap_Exceeded FALSE OR E-stop asserted)
   - DebounceTimer enabled when Gap_Exceeded = TRUE; cleared when
     Gap_Exceeded = FALSE; no same-scan priority issue (TON called
     once with final enable state)
   - Reset: E-stop immediate reset, then return to POWER_UP_INHIBIT
   -----------------------------------------------------------------
   E-STOP PRIORITY (Weld_E_Stop_NC = FALSE):
   - Operator_Alert immediately FALSE (explicit reset per PUB004)
   - Incomplete debounce timing cleared (TON.ET reset via re-call
     with IN=FALSE when E-stop detected)
   - Weld_Soft_Start_Active := FALSE (inhibition cancelled)
   - Same-scan: evaluated before state logic; no race condition
   -----------------------------------------------------------------
   Units/Boundaries:
   - Power-up inhibit: 5s (T#5s), LTIME resolution
   - DebounceTime: caller-supplied TIME, must be positive (PUB003)
   - TON.Q activates at ET >= PT; ET saturates at PT
   - Direction conflicts: not applicable (no axis outputs)
   =================================================================
*)
VAR_INPUT
    Gap_Exceeded: BOOL;
    Weld_E_Stop_NC: BOOL;
    DebounceTime: TIME;
END_VAR

VAR_OUTPUT
    Operator_Alert: BOOL;
    Weld_Soft_Start_Active: BOOL;
END_VAR

VAR
    // Power-up initialization timer: 5-second inhibit period
    PowerUpTimer: TON;
    // Gap signal debounce timer during normal monitoring
    DebounceTimer: TON;
END_VAR

// E-STOP PRIORITY: Immediate deactivation per PUB004
// Evaluated first to ensure same-scan priority over state transitions
IF NOT Weld_E_Stop_NC THEN
    // Operator_Alert immediately FALSE
    Operator_Alert := FALSE;
    // Clear any incomplete debounce timing (re-call with IN=FALSE clears ET)
    DebounceTimer(IN := FALSE, PT := DebounceTime);
    // Cancel power-up inhibition (soft start no longer valid)
    Weld_Soft_Start_Active := FALSE;
    // Restart power-up timer on next rising edge of E-stop release
    PowerUpTimer(IN := FALSE, PT := T#5s);
ELSE
    // E-stop inactive (Weld_E_Stop_NC = TRUE): normal/state logic

    // Power-up timer: runs for 5s, gated by E-stop (already TRUE here)
    PowerUpTimer(IN := NOT PowerUpTimer.Q, PT := T#5s);

    // Determine current operating phase
    IF NOT PowerUpTimer.Q THEN
        // POWER_UP_INHIBIT state: 5-second initialization period
        // PUB001: Operator_Alert = FALSE during inhibit
        Operator_Alert := FALSE;
        // PUB002: Weld_Soft_Start_Active = TRUE during inhibit
        Weld_Soft_Start_Active := TRUE;
        // PUB003: Gap debounce time does NOT accumulate during inhibit
        // Timer not called, so no timing accumulation
    ELSE
        // NORMAL_MONITORING state: after 5-second inhibit completes
        // PUB002: Weld_Soft_Start_Active = FALSE after inhibit
        Weld_Soft_Start_Active := FALSE;

        // Debounce logic: accumulate time only when Gap_Exceeded = TRUE
        // When Gap_Exceeded = FALSE, timer resets (IN=FALSE clears ET)
        DebounceTimer(
            IN := Gap_Exceeded,
            PT := DebounceTime
        );

        // Operator_Alert activated after debounce completes (PUB003)
        // Retention: remains TRUE until Gap_Exceeded FALSE OR E-stop
        Operator_Alert := DebounceTimer.Q;
    END_IF;
END_IF;
END_FUNCTION_BLOCK

(* ---- public-easy-05.raw_candidate_01.st ---- *)
FUNCTION_BLOCK WeldGapAlarm
(* ENGINEERING_CONTRACT
   =================================================================
   States & Retention (outputs per PUB001-PUB006):
   -----------------------------------------------------------------
   State: POWER_UP_INHIBIT (5s after power-up, no E-stop)
   - Weld_Soft_Start_Active := TRUE (activation: power-up entry)
   - Operator_Alert := FALSE (held, no alarm during inhibit)
   - Gap debounce does NOT accumulate (timer gated OFF)
   - Retention: held until 5s elapsed OR E-stop asserted
   -----------------------------------------------------------------
   State: NORMAL_MONITORING (after 5s inhibit, no E-stop)
   - Weld_Soft_Start_Active := FALSE (deactivated, no reset input)
   - Operator_Alert := TRUE only when DebounceTimer.Q = TRUE
     (activation: Gap_Exceeded TRUE for DebounceTime; retention:
      held until Gap_Exceeded FALSE OR E-stop asserted)
   - DebounceTimer enabled when Gap_Exceeded = TRUE; cleared when
     Gap_Exceeded = FALSE; no same-scan priority issue (TON called
     once with final enable state)
   - Reset: E-stop immediate reset, then return to POWER_UP_INHIBIT
   -----------------------------------------------------------------
   E-STOP PRIORITY (Weld_E_Stop_NC = FALSE):
   - Operator_Alert immediately FALSE (explicit reset per PUB004)
   - Incomplete debounce timing cleared (TON.ET reset via re-call
     with IN=FALSE when E-stop detected)
   - Weld_Soft_Start_Active := FALSE (inhibition cancelled)
   - Same-scan: evaluated before state logic; no race condition
   -----------------------------------------------------------------
   Units/Boundaries:
   - Power-up inhibit: 5s (T#5s), LTIME resolution
   - DebounceTime: caller-supplied TIME, must be positive (PUB003)
   - TON.Q activates at ET >= PT; ET saturates at PT
   - Direction conflicts: not applicable (no axis outputs)
   =================================================================
*)
VAR
    // Power-up initialization timer: 5-second inhibit period
    PowerUpTimer: TON;
    // Gap signal debounce timer during normal monitoring
    DebounceTimer: TON;
END_VAR

// E-STOP PRIORITY: Immediate deactivation per PUB004
// Evaluated first to ensure same-scan priority over state transitions
IF NOT Weld_E_Stop_NC THEN
    // Operator_Alert immediately FALSE
    Operator_Alert := FALSE;
    // Clear any incomplete debounce timing (re-call with IN=FALSE clears ET)
    DebounceTimer(IN := FALSE, PT := DebounceTime);
    // Cancel power-up inhibition (soft start no longer valid)
    Weld_Soft_Start_Active := FALSE;
    // Restart power-up timer on next rising edge of E-stop release
    PowerUpTimer(IN := FALSE, PT := T#5s);
ELSE
    // E-stop inactive (Weld_E_Stop_NC = TRUE): normal/state logic

    // Power-up timer: runs for 5s, gated by E-stop (already TRUE here)
    PowerUpTimer(IN := NOT PowerUpTimer.Q, PT := T#5s);

    // Determine current operating phase
    IF NOT PowerUpTimer.Q THEN
        // POWER_UP_INHIBIT state: 5-second initialization period
        // PUB001: Operator_Alert = FALSE during inhibit
        Operator_Alert := FALSE;
        // PUB002: Weld_Soft_Start_Active = TRUE during inhibit
        Weld_Soft_Start_Active := TRUE;
        // PUB003: Gap debounce time does NOT accumulate during inhibit
        // Timer not called, so no timing accumulation
    ELSE
        // NORMAL_MONITORING state: after 5-second inhibit completes
        // PUB002: Weld_Soft_Start_Active = FALSE after inhibit
        Weld_Soft_Start_Active := FALSE;

        // Debounce logic: accumulate time only when Gap_Exceeded = TRUE
        // When Gap_Exceeded = FALSE, timer resets (IN=FALSE clears ET)
        DebounceTimer(
            IN := Gap_Exceeded,
            PT := DebounceTime
        );

        // Operator_Alert activated after debounce completes (PUB003)
        // Retention: remains TRUE until Gap_Exceeded FALSE OR E-stop
        Operator_Alert := DebounceTimer.Q;
    END_IF;
END_IF;
END_FUNCTION_BLOCK

(* ---- public-easy-05.raw_candidate_02.st ---- *)
FUNCTION_BLOCK WeldGapAlarm
(* ENGINEERING_CONTRACT
   =================================================================
   States & Retention (outputs per PUB001-PUB006):
   -----------------------------------------------------------------
   State: POWER_UP_INHIBIT (5s after power-up, no E-stop)
   - Weld_Soft_Start_Active := TRUE (activation: power-up entry)
   - Operator_Alert := FALSE (held, no alarm during inhibit)
   - Gap debounce does NOT accumulate (timer gated OFF)
   - Retention: held until 5s elapsed OR E-stop asserted
   -----------------------------------------------------------------
   State: NORMAL_MONITORING (after 5s inhibit, no E-stop)
   - Weld_Soft_Start_Active := FALSE (deactivated, no reset input)
   - Operator_Alert := TRUE only when DebounceTimer.Q = TRUE
     (activation: Gap_Exceeded TRUE for DebounceTime; retention:
      held until Gap_Exceeded FALSE OR E-stop asserted)
   - DebounceTimer enabled when Gap_Exceeded = TRUE; cleared when
     Gap_Exceeded = FALSE; no same-scan priority issue (TON called
     once with final enable state)
   - Reset: E-stop immediate reset, then return to POWER_UP_INHIBIT
   -----------------------------------------------------------------
   E-STOP PRIORITY (Weld_E_Stop_NC = FALSE):
   - Operator_Alert immediately FALSE (explicit reset per PUB004)
   - Incomplete debounce timing cleared (TON.ET reset via re-call
     with IN=FALSE when E-stop detected)
   - Weld_Soft_Start_Active := FALSE (inhibition cancelled)
   - Same-scan: evaluated before state logic; no race condition
   -----------------------------------------------------------------
   Units/Boundaries:
   - Power-up inhibit: 5s (T#5s), LTIME resolution
   - DebounceTime: caller-supplied TIME, must be positive (PUB003)
   - TON.Q activates at ET >= PT; ET saturates at PT
   - Direction conflicts: not applicable (no axis outputs)
   =================================================================
*)
VAR_INPUT
    Gap_Exceeded: BOOL;
    Weld_E_Stop_NC: BOOL;
    DebounceTime: TIME;
END_VAR

VAR_OUTPUT
    Operator_Alert: BOOL;
    Weld_Soft_Start_Active: BOOL;
END_VAR

VAR
    // Power-up initialization timer: 5-second inhibit period
    PowerUpTimer: TON;
    // Gap signal debounce timer during normal monitoring
    DebounceTimer: TON;
END_VAR

// E-STOP PRIORITY: Immediate deactivation per PUB004
// Evaluated first to ensure same-scan priority over state transitions
IF NOT Weld_E_Stop_NC THEN
    // Operator_Alert immediately FALSE
    Operator_Alert := FALSE;
    // Clear any incomplete debounce timing (re-call with IN=FALSE clears ET)
    DebounceTimer(IN := FALSE, PT := DebounceTime);
    // Cancel power-up inhibition (soft start no longer valid)
    Weld_Soft_Start_Active := FALSE;
    // Restart power-up timer on next rising edge of E-stop release
    PowerUpTimer(IN := FALSE, PT := T#5s);
ELSE
    // E-stop inactive (Weld_E_Stop_NC = TRUE): normal/state logic

    // Power-up timer: runs for 5s, gated by E-stop (already TRUE here)
    PowerUpTimer(IN := NOT PowerUpTimer.Q, PT := T#5s);

    // Determine current operating phase
    IF NOT PowerUpTimer.Q THEN
        // POWER_UP_INHIBIT state: 5-second initialization period
        // PUB001: Operator_Alert = FALSE during inhibit
        Operator_Alert := FALSE;
        // PUB002: Weld_Soft_Start_Active = TRUE during inhibit
        Weld_Soft_Start_Active := TRUE;
        // PUB003: Gap debounce time does NOT accumulate during inhibit
        // Timer not called, so no timing accumulation
    ELSE
        // NORMAL_MONITORING state: after 5-second inhibit completes
        // PUB002: Weld_Soft_Start_Active = FALSE after inhibit
        Weld_Soft_Start_Active := FALSE;

        // Debounce logic: accumulate time only when Gap_Exceeded = TRUE
        // When Gap_Exceeded = FALSE, timer resets (IN=FALSE clears ET)
        DebounceTimer(
            IN := Gap_Exceeded,
            PT := DebounceTime
        );

        // Operator_Alert activated after debounce completes (PUB003)
        // Retention: remains TRUE until Gap_Exceeded FALSE OR E-stop
        Operator_Alert := DebounceTimer.Q;
    END_IF;
END_IF;
END_FUNCTION_BLOCK

(* ---- public-easy-06.candidate_01.st ---- *)
FUNCTION_BLOCK AerationBlowerDelayedStart
(*
    ENGINEERING_CONTRACT
    PUB001: BLOWER_RUN activates only after DO_LOW AND AERATION_E_STOP_NC are TRUE continuously for 5 seconds.
    PUB002: BLOWER_RUN and timer reset immediately when DO_LOW=FALSE OR AERATION_E_STOP_NC=FALSE (no partial credit).
    PUB003: AERATION_BLOWER_CYCLE_COUNT increments on FALSE-to-TRUE (rising) edge of BLOWER_RUN; no repeat during sustained TRUE.
    PUB004: Power-up initializes BLOWER_RUN=FALSE and AERATION_BLOWER_CYCLE_COUNT=0; no prior state retained.
    Activation: BLOWER_RUN = TON.Q (PT=5000ms, IN=DO_LOW AND AERATION_E_STOP_NC).
    Retention: BLOWER_RUN held TRUE while start conditions remain satisfied without stop event.
    Reset/Deactivation: Timer.IN:=FALSE forces TON.Q:=FALSE on same scan as condition loss.
    Same-scan priority: Final condition state determines timer enable before TON call; output assigned after.
    Units/Boundaries: TON PT=TIME#5s (5000ms); threshold is >= PT (TON.Q true when ET >= PT).
*)

VAR_INPUT
    DO_LOW              : BOOL;  (* Dissolved oxygen below threshold; aeration demand *)
    AERATION_E_STOP_NC  : BOOL;  (* TRUE=inactive, FALSE=emergency stop active *)
END_VAR

VAR_OUTPUT
    BLOWER_RUN                  : BOOL;  (* Blower motor run command *)
    AERATION_BLOWER_CYCLE_COUNT : UINT;  (* Count of blower start cycles *)
END_VAR

VAR
    tmp_Rise : R_TRIG;  (* Rising-edge detector for cycle counting *)
    tmp_Ton  : TON;     (* 5-second start delay timer *)
END_VAR

(* Cycle counter rising-edge detector *)
tmp_Rise(CLK := BLOWER_RUN);
IF tmp_Rise.Q THEN
    AERATION_BLOWER_CYCLE_COUNT := AERATION_BLOWER_CYCLE_COUNT + UINT#1;
END_IF;

(* Start-delay timer: IN is TRUE only when both demand present and E-stop inactive *)
tmp_Ton.IN  := DO_LOW AND AERATION_E_STOP_NC;
tmp_Ton.PT  := T#5S;
tmp_Ton();

(* Blower command follows timer completion; both IN and Q go FALSE on same scan when conditions drop *)
BLOWER_RUN := tmp_Ton.Q;

END_FUNCTION_BLOCK

(* CONTRACT_RULES [] *)

(* ---- public-easy-06.patch_base_02.st ---- *)
FUNCTION_BLOCK AerationBlowerDelayedStart
(*
    ENGINEERING_CONTRACT
    PUB001: BLOWER_RUN activates only after DO_LOW AND AERATION_E_STOP_NC are TRUE continuously for 5 seconds.
    PUB002: BLOWER_RUN and timer reset immediately when DO_LOW=FALSE OR AERATION_E_STOP_NC=FALSE (no partial credit).
    PUB003: AERATION_BLOWER_CYCLE_COUNT increments on FALSE-to-TRUE (rising) edge of BLOWER_RUN; no repeat during sustained TRUE.
    PUB004: Power-up initializes BLOWER_RUN=FALSE and AERATION_BLOWER_CYCLE_COUNT=0; no prior state retained.
    Activation: BLOWER_RUN = TON.Q (PT=5000ms, IN=DO_LOW AND AERATION_E_STOP_NC).
    Retention: BLOWER_RUN held TRUE while start conditions remain satisfied without stop event.
    Reset/Deactivation: Timer.IN:=FALSE forces TON.Q:=FALSE on same scan as condition loss.
    Same-scan priority: Final condition state determines timer enable before TON call; output assigned after.
    Units/Boundaries: TON PT=TIME#5s (5000ms); threshold is >= PT (TON.Q true when ET >= PT).
*)

VAR_INPUT
    DO_LOW              : BOOL;  (* Dissolved oxygen below threshold; aeration demand *)
    AERATION_E_STOP_NC  : BOOL;  (* TRUE=inactive, FALSE=emergency stop active *)
END_VAR

VAR_OUTPUT
    BLOWER_RUN                  : BOOL;  (* Blower motor run command *)
    AERATION_BLOWER_CYCLE_COUNT : UINT;  (* Count of blower start cycles *)
END_VAR

VAR
    tmp_Rise : R_TRIG;  (* Rising-edge detector for cycle counting *)
    tmp_Ton  : TON;     (* 5-second start delay timer *)
END_VAR

(* Cycle counter rising-edge detector *)
tmp_Rise(CLK := BLOWER_RUN);
IF tmp_Rise.Q THEN
    AERATION_BLOWER_CYCLE_COUNT := AERATION_BLOWER_CYCLE_COUNT + UINT#1;
END_IF;

(* Start-delay timer: IN is TRUE only when both demand present and E-stop inactive *)
tmp_Ton.IN  := DO_LOW AND AERATION_E_STOP_NC;
tmp_Ton.PT  := T#5S;
tmp_Ton();

(* Blower command follows timer completion; both IN and Q go FALSE on same scan when conditions drop *)
BLOWER_RUN := tmp_Ton.Q;

END_FUNCTION_BLOCK

(* CONTRACT_RULES [] *)

(* ---- public-easy-06.patch_base_03.st ---- *)
FUNCTION_BLOCK AerationBlowerDelayedStart
(*
    ENGINEERING_CONTRACT
    PUB001: BLOWER_RUN activates only after DO_LOW AND AERATION_E_STOP_NC are TRUE continuously for 5 seconds.
    PUB002: BLOWER_RUN and timer reset immediately when DO_LOW=FALSE OR AERATION_E_STOP_NC=FALSE (no partial credit).
    PUB003: AERATION_BLOWER_CYCLE_COUNT increments on FALSE-to-TRUE (rising) edge of BLOWER_RUN; no repeat during sustained TRUE.
    PUB004: Power-up initializes BLOWER_RUN=FALSE and AERATION_BLOWER_CYCLE_COUNT=0; no prior state retained.
    Activation: BLOWER_RUN = TON.Q (PT=5000ms, IN=DO_LOW AND AERATION_E_STOP_NC).
    Retention: BLOWER_RUN held TRUE while start conditions remain satisfied without stop event.
    Reset/Deactivation: Timer.IN:=FALSE forces TON.Q:=FALSE on same scan as condition loss.
    Same-scan priority: Final condition state determines timer enable before TON call; output assigned after.
    Units/Boundaries: TON PT=TIME#5s (5000ms); threshold is >= PT (TON.Q true when ET >= PT).
*)

VAR_INPUT
    DO_LOW              : BOOL;  (* Dissolved oxygen below threshold; aeration demand *)
    AERATION_E_STOP_NC  : BOOL;  (* TRUE=inactive, FALSE=emergency stop active *)
END_VAR

VAR_OUTPUT
    BLOWER_RUN                  : BOOL;  (* Blower motor run command *)
    AERATION_BLOWER_CYCLE_COUNT : UINT;  (* Count of blower start cycles *)
END_VAR

VAR
    tmp_Rise : R_TRIG;  (* Rising-edge detector for cycle counting *)
    tmp_Ton  : TON;     (* 5-second start delay timer *)
END_VAR

(* Cycle counter rising-edge detector *)
tmp_Rise(CLK := BLOWER_RUN);
IF tmp_Rise.Q THEN
    AERATION_BLOWER_CYCLE_COUNT := AERATION_BLOWER_CYCLE_COUNT + UINT#1;
END_IF;

(* Start-delay timer: IN is TRUE only when both demand present and E-stop inactive *)
tmp_Ton.IN  := DO_LOW AND AERATION_E_STOP_NC;
tmp_Ton.PT  := T#5S;
tmp_Ton();

(* Blower command follows timer completion; both IN and Q go FALSE on same scan when conditions drop *)
BLOWER_RUN := tmp_Ton.Q;

END_FUNCTION_BLOCK

(* CONTRACT_RULES [] *)

(* ---- public-easy-06.raw_candidate_01.st ---- *)
FUNCTION_BLOCK AerationBlowerDelayedStart
(*
    ENGINEERING_CONTRACT
    PUB001: BLOWER_RUN activates only after DO_LOW AND AERATION_E_STOP_NC are TRUE continuously for 5 seconds.
    PUB002: BLOWER_RUN and timer reset immediately when DO_LOW=FALSE OR AERATION_E_STOP_NC=FALSE (no partial credit).
    PUB003: AERATION_BLOWER_CYCLE_COUNT increments on FALSE-to-TRUE (rising) edge of BLOWER_RUN; no repeat during sustained TRUE.
    PUB004: Power-up initializes BLOWER_RUN=FALSE and AERATION_BLOWER_CYCLE_COUNT=0; no prior state retained.
    Activation: BLOWER_RUN = TON.Q (PT=5000ms, IN=DO_LOW AND AERATION_E_STOP_NC).
    Retention: BLOWER_RUN held TRUE while start conditions remain satisfied without stop event.
    Reset/Deactivation: Timer.IN:=FALSE forces TON.Q:=FALSE on same scan as condition loss.
    Same-scan priority: Final condition state determines timer enable before TON call; output assigned after.
    Units/Boundaries: TON PT=TIME#5s (5000ms); threshold is >= PT (TON.Q true when ET >= PT).
*)

VAR_INPUT
    DO_LOW              : BOOL;  (* Dissolved oxygen below threshold; aeration demand *)
    AERATION_E_STOP_NC  : BOOL;  (* TRUE=inactive, FALSE=emergency stop active *)
END_VAR

VAR_OUTPUT
    BLOWER_RUN                  : BOOL;  (* Blower motor run command *)
    AERATION_BLOWER_CYCLE_COUNT : UINT;  (* Count of blower start cycles *)
END_VAR

VAR
    tmp_Rise : R_TRIG;  (* Rising-edge detector for cycle counting *)
    tmp_Ton  : TON;     (* 5-second start delay timer *)
END_VAR

(* Cycle counter rising-edge detector *)
tmp_Rise(CLK := BLOWER_RUN);
IF tmp_Rise.Q THEN
    AERATION_BLOWER_CYCLE_COUNT := AERATION_BLOWER_CYCLE_COUNT + UINT#1;
END_IF;

(* Start-delay timer: IN is TRUE only when both demand present and E-stop inactive *)
tmp_Ton.IN  := DO_LOW AND AERATION_E_STOP_NC;
tmp_Ton.PT  := T#5S;
tmp_Ton();

(* Blower command follows timer completion; both IN and Q go FALSE on same scan when conditions drop *)
BLOWER_RUN := tmp_Ton.Q;

END_FUNCTION_BLOCK

(* CONTRACT_RULES [] *)

(* ---- public-hard-03.candidate_01.st ---- *)
FUNCTION_BLOCK FB_RecipeManager
VAR_INPUT
    addRecipe      : BOOL;
    deleteRecipe   : BOOL;
    modifyRecipe   : BOOL;
    queryRecipe    : BOOL;
    recipeIn       : ST_Recipe;
END_VAR

VAR_OUTPUT
    recipeAdded        : BOOL;
    recipeDeleted      : BOOL;
    recipeModified     : BOOL;
    recipeQueryResult  : ST_Recipe;
    error              : BOOL;
    status             : WORD;
END_VAR

VAR_IN_OUT
    recipe : ARRAY[1..10] OF ST_Recipe;
END_VAR

VAR
    tmp_foundIndex : INT;
    tmp_emptyIndex : INT;
    tmp_i          : INT;
END_VAR

(*
ENGINEERING_CONTRACT
===================
Operation sequencing (PUB001-PUB005, PUB007-PUB012):
- Commands evaluated in priority order: DELETE > ADD > MODIFY > QUERY when multiple asserted.
- All success pulses are same-scan; no retention across scans.

Query (PUB008):
  Activation:    queryRecipe rising edge or held high during scan.
  Retention:     recipeQueryResult valid until next scan or successful QUERY.
  Reset:         error and status cleared at start of scan.
  Error codes:   16#8001 = recipe not found.
  Units:         Status WORD error code.

Add (PUB009):
  Activation:    addRecipe rising edge or held high.
  Retention:     Stored in smallest-index empty slot; persists until delete.
  Reset:         None (persistent storage).
  Error codes:   16#8002 = duplicate ID; 16#8003 = database full.
  Same-scan:     Duplicate check before empty-slot check.

Delete (PUB010):
  Activation:    deleteRecipe rising edge or held high.
  Retention:     recipeID forced to 0 (empty slot marker).
  Reset:         Implicit (setting ID to 0 removes it).
  Error codes:   16#8004 = recipe not found.

Modify (PUB011-PUB012):
  Activation:    modifyRecipe rising edge or held high.
  Retention:     Full recipe replacement at found slot.
  Reset:         None.
  Error codes:   16#8005 = recipe not found.
*)

(* CONTRACT_RULES [] *)

tmp_foundIndex := 0;
tmp_emptyIndex := 0;
error := FALSE;
status := 16#0;
recipeAdded := FALSE;
recipeDeleted := FALSE;
recipeModified := FALSE;

IF deleteRecipe THEN
    tmp_foundIndex := 0;
    FOR tmp_i := 1 TO 10 DO
        IF recipe[tmp_i].recipeID <> 0 AND recipe[tmp_i].recipeID = recipeIn.recipeID THEN
            tmp_foundIndex := tmp_i;
            EXIT;
        END_IF;
    END_FOR;

    IF tmp_foundIndex = 0 THEN
        error := TRUE;
        status := 16#8004;
    ELSE
        recipe[tmp_foundIndex].recipeID := 0;
        recipeDeleted := TRUE;
    END_IF;

ELSIF addRecipe THEN
    tmp_foundIndex := 0;
    tmp_emptyIndex := 0;

    FOR tmp_i := 1 TO 10 DO
        IF recipe[tmp_i].recipeID <> 0 AND recipe[tmp_i].recipeID = recipeIn.recipeID THEN
            tmp_foundIndex := tmp_i;
            EXIT;
        END_IF;
    END_FOR;

    IF tmp_foundIndex <> 0 THEN
        error := TRUE;
        status := 16#8002;
    ELSE
        FOR tmp_i := 1 TO 10 DO
            IF recipe[tmp_i].recipeID = 0 AND tmp_emptyIndex = 0 THEN
                tmp_emptyIndex := tmp_i;
                EXIT;
            END_IF;
        END_FOR;

        IF tmp_emptyIndex = 0 THEN
            error := TRUE;
            status := 16#8003;
        ELSE
            recipe[tmp_emptyIndex] := recipeIn;
            recipeAdded := TRUE;
        END_IF;
    END_IF;

ELSIF modifyRecipe THEN
    tmp_foundIndex := 0;
    FOR tmp_i := 1 TO 10 DO
        IF recipe[tmp_i].recipeID <> 0 AND recipe[tmp_i].recipeID = recipeIn.recipeID THEN
            tmp_foundIndex := tmp_i;
            EXIT;
        END_IF;
    END_FOR;

    IF tmp_foundIndex = 0 THEN
        error := TRUE;
        status := 16#8005;
    ELSE
        recipe[tmp_foundIndex] := recipeIn;
        recipeModified := TRUE;
    END_IF;

ELSIF queryRecipe THEN
    tmp_foundIndex := 0;
    FOR tmp_i := 1 TO 10 DO
        IF recipe[tmp_i].recipeID <> 0 AND recipe[tmp_i].recipeID = recipeIn.recipeID THEN
            tmp_foundIndex := tmp_i;
            EXIT;
        END_IF;
    END_FOR;

    IF tmp_foundIndex = 0 THEN
        error := TRUE;
        status := 16#8001;
    ELSE
        recipeQueryResult := recipe[tmp_foundIndex];
    END_IF;
END_IF;

END_FUNCTION_BLOCK

(* ---- public-hard-03.candidate_02.st ---- *)
TYPE ST_Recipe :
STRUCT
    recipeID               : INT;
    ingredientType         : INT;
    ingredientRatio        : REAL;
    productionTemperature  : REAL;
END_STRUCT
END_TYPE;

FUNCTION_BLOCK FB_RecipeManager
VAR_INPUT
    addRecipe      : BOOL;
    deleteRecipe   : BOOL;
    modifyRecipe   : BOOL;
    queryRecipe    : BOOL;
    recipeIn       : ST_Recipe;
END_VAR

VAR_OUTPUT
    recipeAdded        : BOOL;
    recipeDeleted      : BOOL;
    recipeModified     : BOOL;
    recipeQueryResult  : ST_Recipe;
    error              : BOOL;
    status             : WORD;
END_VAR

VAR_IN_OUT
    recipe : ARRAY[1..10] OF ST_Recipe;
END_VAR

VAR
    tmp_foundIndex : INT;
    tmp_emptyIndex : INT;
    tmp_i          : INT;
END_VAR

(*
ENGINEERING_CONTRACT
===================
Operation sequencing (PUB001-PUB005, PUB007-PUB012):
- Commands evaluated in priority order: DELETE > ADD > MODIFY > QUERY when multiple asserted.
- All success pulses are same-scan; no retention across scans.

Query (PUB008):
  Activation:    queryRecipe rising edge or held high during scan.
  Retention:     recipeQueryResult valid until next scan or successful QUERY.
  Reset:         error and status cleared at start of scan.
  Error codes:   16#8001 = recipe not found.
  Units:         Status WORD error code.

Add (PUB009):
  Activation:    addRecipe rising edge or held high.
  Retention:     Stored in smallest-index empty slot; persists until delete.
  Reset:         None (persistent storage).
  Error codes:   16#8002 = duplicate ID; 16#8003 = database full.
  Same-scan:     Duplicate check before empty-slot check.

Delete (PUB010):
  Activation:    deleteRecipe rising edge or held high.
  Retention:     recipeID forced to 0 (empty slot marker).
  Reset:         Implicit (setting ID to 0 removes it).
  Error codes:   16#8004 = recipe not found.

Modify (PUB011-PUB012):
  Activation:    modifyRecipe rising edge or held high.
  Retention:     Full recipe replacement at found slot.
  Reset:         None.
  Error codes:   16#8005 = recipe not found.
*)

(* CONTRACT_RULES [] *)

tmp_foundIndex := 0;
tmp_emptyIndex := 0;
error := FALSE;
status := 16#0;
recipeAdded := FALSE;
recipeDeleted := FALSE;
recipeModified := FALSE;

IF deleteRecipe THEN
    tmp_foundIndex := 0;
    FOR tmp_i := 1 TO 10 DO
        IF recipe[tmp_i].recipeID <> 0 AND recipe[tmp_i].recipeID = recipeIn.recipeID THEN
            tmp_foundIndex := tmp_i;
            EXIT;
        END_IF;
    END_FOR;

    IF tmp_foundIndex = 0 THEN
        error := TRUE;
        status := 16#8004;
    ELSE
        recipe[tmp_foundIndex].recipeID := 0;
        recipeDeleted := TRUE;
    END_IF;

ELSIF addRecipe THEN
    tmp_foundIndex := 0;
    tmp_emptyIndex := 0;

    FOR tmp_i := 1 TO 10 DO
        IF recipe[tmp_i].recipeID <> 0 AND recipe[tmp_i].recipeID = recipeIn.recipeID THEN
            tmp_foundIndex := tmp_i;
            EXIT;
        END_IF;
    END_FOR;

    IF tmp_foundIndex <> 0 THEN
        error := TRUE;
        status := 16#8002;
    ELSE
        FOR tmp_i := 1 TO 10 DO
            IF recipe[tmp_i].recipeID = 0 AND tmp_emptyIndex = 0 THEN
                tmp_emptyIndex := tmp_i;
                EXIT;
            END_IF;
        END_FOR;

        IF tmp_emptyIndex = 0 THEN
            error := TRUE;
            status := 16#8003;
        ELSE
            recipe[tmp_emptyIndex] := recipeIn;
            recipeAdded := TRUE;
        END_IF;
    END_IF;

ELSIF modifyRecipe THEN
    tmp_foundIndex := 0;
    FOR tmp_i := 1 TO 10 DO
        IF recipe[tmp_i].recipeID <> 0 AND recipe[tmp_i].recipeID = recipeIn.recipeID THEN
            tmp_foundIndex := tmp_i;
            EXIT;
        END_IF;
    END_FOR;

    IF tmp_foundIndex = 0 THEN
        error := TRUE;
        status := 16#8005;
    ELSE
        recipe[tmp_foundIndex] := recipeIn;
        recipeModified := TRUE;
    END_IF;

ELSIF queryRecipe THEN
    tmp_foundIndex := 0;
    FOR tmp_i := 1 TO 10 DO
        IF recipe[tmp_i].recipeID <> 0 AND recipe[tmp_i].recipeID = recipeIn.recipeID THEN
            tmp_foundIndex := tmp_i;
            EXIT;
        END_IF;
    END_FOR;

    IF tmp_foundIndex = 0 THEN
        error := TRUE;
        status := 16#8001;
    ELSE
        recipeQueryResult := recipe[tmp_foundIndex];
    END_IF;
END_IF;

END_FUNCTION_BLOCK

(* ---- public-hard-03.patch_base_02.st ---- *)
FUNCTION_BLOCK FB_RecipeManager
VAR_INPUT
    addRecipe      : BOOL;
    deleteRecipe   : BOOL;
    modifyRecipe   : BOOL;
    queryRecipe    : BOOL;
    recipeIn       : ST_Recipe;
END_VAR

VAR_OUTPUT
    recipeAdded        : BOOL;
    recipeDeleted      : BOOL;
    recipeModified     : BOOL;
    recipeQueryResult  : ST_Recipe;
    error              : BOOL;
    status             : WORD;
END_VAR

VAR_IN_OUT
    recipe : ARRAY[1..10] OF ST_Recipe;
END_VAR

VAR
    tmp_foundIndex : INT;
    tmp_emptyIndex : INT;
    tmp_i          : INT;
END_VAR

(*
ENGINEERING_CONTRACT
===================
Operation sequencing (PUB001-PUB005, PUB007-PUB012):
- Commands evaluated in priority order: DELETE > ADD > MODIFY > QUERY when multiple asserted.
- All success pulses are same-scan; no retention across scans.

Query (PUB008):
  Activation:    queryRecipe rising edge or held high during scan.
  Retention:     recipeQueryResult valid until next scan or successful QUERY.
  Reset:         error and status cleared at start of scan.
  Error codes:   16#8001 = recipe not found.
  Units:         Status WORD error code.

Add (PUB009):
  Activation:    addRecipe rising edge or held high.
  Retention:     Stored in smallest-index empty slot; persists until delete.
  Reset:         None (persistent storage).
  Error codes:   16#8002 = duplicate ID; 16#8003 = database full.
  Same-scan:     Duplicate check before empty-slot check.

Delete (PUB010):
  Activation:    deleteRecipe rising edge or held high.
  Retention:     recipeID forced to 0 (empty slot marker).
  Reset:         Implicit (setting ID to 0 removes it).
  Error codes:   16#8004 = recipe not found.

Modify (PUB011-PUB012):
  Activation:    modifyRecipe rising edge or held high.
  Retention:     Full recipe replacement at found slot.
  Reset:         None.
  Error codes:   16#8005 = recipe not found.
*)

(* CONTRACT_RULES [] *)

tmp_foundIndex := 0;
tmp_emptyIndex := 0;
error := FALSE;
status := 16#0;
recipeAdded := FALSE;
recipeDeleted := FALSE;
recipeModified := FALSE;

IF deleteRecipe THEN
    tmp_foundIndex := 0;
    FOR tmp_i := 1 TO 10 DO
        IF recipe[tmp_i].recipeID <> 0 AND recipe[tmp_i].recipeID = recipeIn.recipeID THEN
            tmp_foundIndex := tmp_i;
            EXIT;
        END_IF;
    END_FOR;

    IF tmp_foundIndex = 0 THEN
        error := TRUE;
        status := 16#8004;
    ELSE
        recipe[tmp_foundIndex].recipeID := 0;
        recipeDeleted := TRUE;
    END_IF;

ELSIF addRecipe THEN
    tmp_foundIndex := 0;
    tmp_emptyIndex := 0;

    FOR tmp_i := 1 TO 10 DO
        IF recipe[tmp_i].recipeID <> 0 AND recipe[tmp_i].recipeID = recipeIn.recipeID THEN
            tmp_foundIndex := tmp_i;
            EXIT;
        END_IF;
    END_FOR;

    IF tmp_foundIndex <> 0 THEN
        error := TRUE;
        status := 16#8002;
    ELSE
        FOR tmp_i := 1 TO 10 DO
            IF recipe[tmp_i].recipeID = 0 AND tmp_emptyIndex = 0 THEN
                tmp_emptyIndex := tmp_i;
                EXIT;
            END_IF;
        END_FOR;

        IF tmp_emptyIndex = 0 THEN
            error := TRUE;
            status := 16#8003;
        ELSE
            recipe[tmp_emptyIndex] := recipeIn;
            recipeAdded := TRUE;
        END_IF;
    END_IF;

ELSIF modifyRecipe THEN
    tmp_foundIndex := 0;
    FOR tmp_i := 1 TO 10 DO
        IF recipe[tmp_i].recipeID <> 0 AND recipe[tmp_i].recipeID = recipeIn.recipeID THEN
            tmp_foundIndex := tmp_i;
            EXIT;
        END_IF;
    END_FOR;

    IF tmp_foundIndex = 0 THEN
        error := TRUE;
        status := 16#8005;
    ELSE
        recipe[tmp_foundIndex] := recipeIn;
        recipeModified := TRUE;
    END_IF;

ELSIF queryRecipe THEN
    tmp_foundIndex := 0;
    FOR tmp_i := 1 TO 10 DO
        IF recipe[tmp_i].recipeID <> 0 AND recipe[tmp_i].recipeID = recipeIn.recipeID THEN
            tmp_foundIndex := tmp_i;
            EXIT;
        END_IF;
    END_FOR;

    IF tmp_foundIndex = 0 THEN
        error := TRUE;
        status := 16#8001;
    ELSE
        recipeQueryResult := recipe[tmp_foundIndex];
    END_IF;
END_IF;

END_FUNCTION_BLOCK

(* ---- public-hard-03.patch_base_03.st ---- *)
TYPE ST_Recipe :
STRUCT
    recipeID               : INT;
    ingredientType         : INT;
    ingredientRatio        : REAL;
    productionTemperature  : REAL;
END_STRUCT
END_TYPE;

FUNCTION_BLOCK FB_RecipeManager
VAR_INPUT
    addRecipe      : BOOL;
    deleteRecipe   : BOOL;
    modifyRecipe   : BOOL;
    queryRecipe    : BOOL;
    recipeIn       : ST_Recipe;
END_VAR

VAR_OUTPUT
    recipeAdded        : BOOL;
    recipeDeleted      : BOOL;
    recipeModified     : BOOL;
    recipeQueryResult  : ST_Recipe;
    error              : BOOL;
    status             : WORD;
END_VAR

VAR_IN_OUT
    recipe : ARRAY[1..10] OF ST_Recipe;
END_VAR

VAR
    tmp_foundIndex : INT;
    tmp_emptyIndex : INT;
    tmp_i          : INT;
END_VAR

(*
ENGINEERING_CONTRACT
===================
Operation sequencing (PUB001-PUB005, PUB007-PUB012):
- Commands evaluated in priority order: DELETE > ADD > MODIFY > QUERY when multiple asserted.
- All success pulses are same-scan; no retention across scans.

Query (PUB008):
  Activation:    queryRecipe rising edge or held high during scan.
  Retention:     recipeQueryResult valid until next scan or successful QUERY.
  Reset:         error and status cleared at start of scan.
  Error codes:   16#8001 = recipe not found.
  Units:         Status WORD error code.

Add (PUB009):
  Activation:    addRecipe rising edge or held high.
  Retention:     Stored in smallest-index empty slot; persists until delete.
  Reset:         None (persistent storage).
  Error codes:   16#8002 = duplicate ID; 16#8003 = database full.
  Same-scan:     Duplicate check before empty-slot check.

Delete (PUB010):
  Activation:    deleteRecipe rising edge or held high.
  Retention:     recipeID forced to 0 (empty slot marker).
  Reset:         Implicit (setting ID to 0 removes it).
  Error codes:   16#8004 = recipe not found.

Modify (PUB011-PUB012):
  Activation:    modifyRecipe rising edge or held high.
  Retention:     Full recipe replacement at found slot.
  Reset:         None.
  Error codes:   16#8005 = recipe not found.
*)

(* CONTRACT_RULES [] *)

tmp_foundIndex := 0;
tmp_emptyIndex := 0;
error := FALSE;
status := 16#0;
recipeAdded := FALSE;
recipeDeleted := FALSE;
recipeModified := FALSE;

IF deleteRecipe THEN
    tmp_foundIndex := 0;
    FOR tmp_i := 1 TO 10 DO
        IF recipe[tmp_i].recipeID <> 0 AND recipe[tmp_i].recipeID = recipeIn.recipeID THEN
            tmp_foundIndex := tmp_i;
            EXIT;
        END_IF;
    END_FOR;

    IF tmp_foundIndex = 0 THEN
        error := TRUE;
        status := 16#8004;
    ELSE
        recipe[tmp_foundIndex].recipeID := 0;
        recipeDeleted := TRUE;
    END_IF;

ELSIF addRecipe THEN
    tmp_foundIndex := 0;
    tmp_emptyIndex := 0;

    FOR tmp_i := 1 TO 10 DO
        IF recipe[tmp_i].recipeID <> 0 AND recipe[tmp_i].recipeID = recipeIn.recipeID THEN
            tmp_foundIndex := tmp_i;
            EXIT;
        END_IF;
    END_FOR;

    IF tmp_foundIndex <> 0 THEN
        error := TRUE;
        status := 16#8002;
    ELSE
        FOR tmp_i := 1 TO 10 DO
            IF recipe[tmp_i].recipeID = 0 AND tmp_emptyIndex = 0 THEN
                tmp_emptyIndex := tmp_i;
                EXIT;
            END_IF;
        END_FOR;

        IF tmp_emptyIndex = 0 THEN
            error := TRUE;
            status := 16#8003;
        ELSE
            recipe[tmp_emptyIndex] := recipeIn;
            recipeAdded := TRUE;
        END_IF;
    END_IF;

ELSIF modifyRecipe THEN
    tmp_foundIndex := 0;
    FOR tmp_i := 1 TO 10 DO
        IF recipe[tmp_i].recipeID <> 0 AND recipe[tmp_i].recipeID = recipeIn.recipeID THEN
            tmp_foundIndex := tmp_i;
            EXIT;
        END_IF;
    END_FOR;

    IF tmp_foundIndex = 0 THEN
        error := TRUE;
        status := 16#8005;
    ELSE
        recipe[tmp_foundIndex] := recipeIn;
        recipeModified := TRUE;
    END_IF;

ELSIF queryRecipe THEN
    tmp_foundIndex := 0;
    FOR tmp_i := 1 TO 10 DO
        IF recipe[tmp_i].recipeID <> 0 AND recipe[tmp_i].recipeID = recipeIn.recipeID THEN
            tmp_foundIndex := tmp_i;
            EXIT;
        END_IF;
    END_FOR;

    IF tmp_foundIndex = 0 THEN
        error := TRUE;
        status := 16#8001;
    ELSE
        recipeQueryResult := recipe[tmp_foundIndex];
    END_IF;
END_IF;

END_FUNCTION_BLOCK

(* ---- public-hard-03.patch_base_04.st ---- *)
TYPE ST_Recipe :
STRUCT
    recipeID               : INT;
    ingredientType         : INT;
    ingredientRatio        : REAL;
    productionTemperature  : REAL;
END_STRUCT
END_TYPE;

FUNCTION_BLOCK FB_RecipeManager
VAR_INPUT
    addRecipe      : BOOL;
    deleteRecipe   : BOOL;
    modifyRecipe   : BOOL;
    queryRecipe    : BOOL;
    recipeIn       : ST_Recipe;
END_VAR

VAR_OUTPUT
    recipeAdded        : BOOL;
    recipeDeleted      : BOOL;
    recipeModified     : BOOL;
    recipeQueryResult  : ST_Recipe;
    error              : BOOL;
    status             : WORD;
END_VAR

VAR_IN_OUT
    recipe : ARRAY[1..10] OF ST_Recipe;
END_VAR

VAR
    tmp_foundIndex : INT;
    tmp_emptyIndex : INT;
    tmp_i          : INT;
END_VAR

(*
ENGINEERING_CONTRACT
===================
Operation sequencing (PUB001-PUB005, PUB007-PUB012):
- Commands evaluated in priority order: DELETE > ADD > MODIFY > QUERY when multiple asserted.
- All success pulses are same-scan; no retention across scans.

Query (PUB008):
  Activation:    queryRecipe rising edge or held high during scan.
  Retention:     recipeQueryResult valid until next scan or successful QUERY.
  Reset:         error and status cleared at start of scan.
  Error codes:   16#8001 = recipe not found.
  Units:         Status WORD error code.

Add (PUB009):
  Activation:    addRecipe rising edge or held high.
  Retention:     Stored in smallest-index empty slot; persists until delete.
  Reset:         None (persistent storage).
  Error codes:   16#8002 = duplicate ID; 16#8003 = database full.
  Same-scan:     Duplicate check before empty-slot check.

Delete (PUB010):
  Activation:    deleteRecipe rising edge or held high.
  Retention:     recipeID forced to 0 (empty slot marker).
  Reset:         Implicit (setting ID to 0 removes it).
  Error codes:   16#8004 = recipe not found.

Modify (PUB011-PUB012):
  Activation:    modifyRecipe rising edge or held high.
  Retention:     Full recipe replacement at found slot.
  Reset:         None.
  Error codes:   16#8005 = recipe not found.
*)

(* CONTRACT_RULES [] *)

tmp_foundIndex := 0;
tmp_emptyIndex := 0;
error := FALSE;
status := 16#0;
recipeAdded := FALSE;
recipeDeleted := FALSE;
recipeModified := FALSE;

IF deleteRecipe THEN
    tmp_foundIndex := 0;
    FOR tmp_i := 1 TO 10 DO
        IF recipe[tmp_i].recipeID <> 0 AND recipe[tmp_i].recipeID = recipeIn.recipeID THEN
            tmp_foundIndex := tmp_i;
            EXIT;
        END_IF;
    END_FOR;

    IF tmp_foundIndex = 0 THEN
        error := TRUE;
        status := 16#8004;
    ELSE
        recipe[tmp_foundIndex].recipeID := 0;
        recipeDeleted := TRUE;
    END_IF;

ELSIF addRecipe THEN
    tmp_foundIndex := 0;
    tmp_emptyIndex := 0;

    FOR tmp_i := 1 TO 10 DO
        IF recipe[tmp_i].recipeID <> 0 AND recipe[tmp_i].recipeID = recipeIn.recipeID THEN
            tmp_foundIndex := tmp_i;
            EXIT;
        END_IF;
    END_FOR;

    IF tmp_foundIndex <> 0 THEN
        error := TRUE;
        status := 16#8002;
    ELSE
        FOR tmp_i := 1 TO 10 DO
            IF recipe[tmp_i].recipeID = 0 AND tmp_emptyIndex = 0 THEN
                tmp_emptyIndex := tmp_i;
                EXIT;
            END_IF;
        END_FOR;

        IF tmp_emptyIndex = 0 THEN
            error := TRUE;
            status := 16#8003;
        ELSE
            recipe[tmp_emptyIndex] := recipeIn;
            recipeAdded := TRUE;
        END_IF;
    END_IF;

ELSIF modifyRecipe THEN
    tmp_foundIndex := 0;
    FOR tmp_i := 1 TO 10 DO
        IF recipe[tmp_i].recipeID <> 0 AND recipe[tmp_i].recipeID = recipeIn.recipeID THEN
            tmp_foundIndex := tmp_i;
            EXIT;
        END_IF;
    END_FOR;

    IF tmp_foundIndex = 0 THEN
        error := TRUE;
        status := 16#8005;
    ELSE
        recipe[tmp_foundIndex] := recipeIn;
        recipeModified := TRUE;
    END_IF;

ELSIF queryRecipe THEN
    tmp_foundIndex := 0;
    FOR tmp_i := 1 TO 10 DO
        IF recipe[tmp_i].recipeID <> 0 AND recipe[tmp_i].recipeID = recipeIn.recipeID THEN
            tmp_foundIndex := tmp_i;
            EXIT;
        END_IF;
    END_FOR;

    IF tmp_foundIndex = 0 THEN
        error := TRUE;
        status := 16#8001;
    ELSE
        recipeQueryResult := recipe[tmp_foundIndex];
    END_IF;
END_IF;

END_FUNCTION_BLOCK
